(* IEC 61131-3 sources: TetherPLC/compat/tc2 (part 5) *)

(* ---- tc2_nci.st ---- *)
// Tc2_NCI — TwinCAT NC-I (TF5100) channel-interpolation surface over
// the builtin FB_MotionAxis (tplc-motion service). This file
// implements the interpolation core: coordinated multi-axis
// setpoint streaming in CyclicSyncPosition (CSP, mode 8).
//
// Model: TwinCAT's NC-I runs a G-code / FIFO interpreter in the NC
// kernel that emits per-axis position setpoints every NC cycle to
// axes in CSP mode. The compat model collapses one in-flight
// geometric block into each FB: FB_NciLine parameterizes a straight
// line across a 3-axis group, advances the path parameter s by
// Velocity*CycleUs each scan, and streams per-axis targets
// (0x607A) with the axes in CSP mode — which is exactly how the NC
// kernel drives CSP axes. There is no backend group registry, so a
// "3D group" is just the X/Y/Z axis handles passed to the block
// (TwinCAT's CfgBuild3DGroup maps to passing those handles).
//
// Time base: the FB has no access to the host clock, so the caller
// supplies the scan period via CycleUs (microseconds); path
// Velocity is then in user-units/second and s += Velocity*CycleUs/1e6
// per scan. Positions/velocities are the backend's int32 user
// units (TwinCAT LREAL — documented gap). Determinism: under --sim,
// CycleUs = step_us makes the path advance a fixed amount per step,
// and CSP snaps each axis to the streamed target so commanded and
// actual positions match.
//
// G-code interpretation lives in Tether: tether_io_motion_server
// exposes an nc.* channel that compiles program text with its G-code
// interpreter, time-parameterizes it with the motion planner (corner
// blending, jerk-limited profiles), and streams CSP setpoints to the
// drives on the mc.time clock. The FB_NciChan blocks below are the
// PLC-side control surface for that channel (TwinCAT Itp* shape);
// there is no in-process interpreter — with no TPLC_MOTION_IO
// endpoint the blocks report the service as unavailable.
//
// Honest gaps: FB_NciLine is the foundational interpreter-free path
// (single block, no queue); the nc.* channel has no PLC-visible
// M-function handshake, R-parameters, zero-shift, or cyclic-channel
// offset tables yet. See DECISIONS D-IMPL-56.
// SPDX-License-Identifier: Apache-2.0 OR MPL-2.0

// ---- F_NciSqrt: Newton (Babylonian) square root for LREAL ----
// The ST layer has no SQRT builtin, so the path length is computed
// with a fixed-iteration Newton iteration. r0 = x/2 + 1 converges
// monotonically for x >= 0; 48 iterations is enough for the full
// int32 path range and keeps the result deterministic.
FUNCTION F_NciSqrt : LREAL
VAR_INPUT
    x : LREAL;
END_VAR
VAR
    r : LREAL;
    k : INT;
END_VAR
    IF x <= 0.0 THEN
        F_NciSqrt := 0.0;
    ELSE
        r := x * 0.5 + 1.0;
        k := 0;
        REPEAT
            r := 0.5 * (r + x / r);
            k := k + 1;
        UNTIL k >= 48
        END_REPEAT;
        F_NciSqrt := r;
    END_IF;
END_FUNCTION

// ---- FB_NciLine: coordinated 3-axis linear move (CSP stream) ----
// On Execute, latches each axis's actual position as the segment
// start, computes deltas and the Euclidean path length, switches
// all three axes to CSP mode, then each scan advances s toward len
// and writes each axis's interpolated TargetPosition. Done when
// s reaches len (all axes arrive simultaneously — a straight line).
// Releasing Execute mid-move aborts: streaming stops, so each axis
// holds its last streamed target (CommandAborted pulses).
FUNCTION_BLOCK FB_NciLine
VAR_INPUT
    Execute : BOOL;
    PosX : DINT;
    PosY : DINT;
    PosZ : DINT;
    Velocity : DINT;    // resultant path velocity, user-units/sec
    CycleUs : DINT;     // scan period, microseconds
    AxisX : UDINT;
    AxisY : UDINT;
    AxisZ : UDINT;
END_VAR
VAR_OUTPUT
    Done : BOOL;
    Busy : BOOL;
    CommandAborted : BOOL;
    Error : BOOL;
    ErrorID : UDINT;
    ActPosX : DINT;     // interpolated commanded positions
    ActPosY : DINT;
    ActPosZ : DINT;
    PathLen : DINT;     // Euclidean path length (user units)
    PathS : DINT;       // current path parameter along the line
END_VAR
VAR
    axX : FB_MotionAxis;
    axY : FB_MotionAxis;
    axZ : FB_MotionAxis;
    exPrev : BOOL;
    exEdge : BOOL;
    active : BOOL;
    sxr : LREAL;
    syr : LREAL;
    szr : LREAL;
    dxr : LREAL;
    dyr : LREAL;
    dzr : LREAL;
    len : LREAL;
    s : LREAL;
    dt : LREAL;
    vel : LREAL;
END_VAR
    // advance every axis's dynamics once per scan (one poll advances
    // the whole pool); bind each instance to its group axis
    axX.OP := 3; axX();
    axX.AXIS := AxisX; axY.AXIS := AxisY; axZ.AXIS := AxisZ;
    exEdge := Execute AND NOT exPrev;
    exPrev := Execute;
    Done := FALSE;
    CommandAborted := FALSE;
    Error := FALSE;
    ErrorID := 0;

    IF exEdge THEN
        // latch the segment start = current actual positions
        axX.OP := 4; axX.INDEX := 16#6064; axX();
        sxr := DINT_TO_LREAL(axX.VALUE);
        axY.OP := 4; axY.INDEX := 16#6064; axY();
        syr := DINT_TO_LREAL(axY.VALUE);
        axZ.OP := 4; axZ.INDEX := 16#6064; axZ();
        szr := DINT_TO_LREAL(axZ.VALUE);
        dxr := DINT_TO_LREAL(PosX) - sxr;
        dyr := DINT_TO_LREAL(PosY) - syr;
        dzr := DINT_TO_LREAL(PosZ) - szr;
        len := F_NciSqrt(dxr * dxr + dyr * dyr + dzr * dzr);
        PathLen := TRUNC(len);
        dt := DINT_TO_LREAL(CycleUs) / 1000000.0;
        vel := DINT_TO_LREAL(Velocity);
        s := 0.0;
        IF len < 0.5 THEN
            // already at the target — nothing to stream
            active := FALSE;
            Done := TRUE;
        ELSE
            // put the group into CyclicSyncPosition (mode 8)
            axX.OP := 5; axX.INDEX := 16#6060; axX.VALUE := 8; axX();
            axY.OP := 5; axY.INDEX := 16#6060; axY.VALUE := 8; axY();
            axZ.OP := 5; axZ.INDEX := 16#6060; axZ.VALUE := 8; axZ();
            active := TRUE;
        END_IF;
    END_IF;

    IF active THEN
        IF Execute THEN
            // advance the path parameter and clamp at the end
            s := s + vel * dt;
            IF s >= len THEN
                s := len;
                active := FALSE;
                Done := TRUE;
            END_IF;
            PathS := TRUNC(s);
            // stream the interpolated setpoints to each CSP axis
            ActPosX := TRUNC(sxr + dxr * s / len);
            ActPosY := TRUNC(syr + dyr * s / len);
            ActPosZ := TRUNC(szr + dzr * s / len);
            axX.OP := 5; axX.INDEX := 16#607A; axX.VALUE := ActPosX; axX();
            axY.OP := 5; axY.INDEX := 16#607A; axY.VALUE := ActPosY; axY();
            axZ.OP := 5; axZ.INDEX := 16#607A; axZ.VALUE := ActPosZ; axZ();
        ELSE
            // aborted: stop streaming so each axis holds its last
            // CSP setpoint (position freezes in place)
            active := FALSE;
            CommandAborted := TRUE;
        END_IF;
    END_IF;
    Busy := active;
END_FUNCTION_BLOCK

// ---- FB_NciEStop: cut power to a 3-axis group ----
// On Execute it writes DisableVoltage (controlword 0x0000) to each
// axis so the group coasts to a stop; Status reports all three
// axes left OperationEnabled. Honest E-stop: a real NC fault also
// freezes the interpolator, which the caller models by releasing
// FB_NciLine's Execute.
FUNCTION_BLOCK FB_NciEStop
VAR_INPUT
    Execute : BOOL;
    AxisX : UDINT;
    AxisY : UDINT;
    AxisZ : UDINT;
END_VAR
VAR_OUTPUT
    Status : BOOL;
    Busy : BOOL;
    Error : BOOL;
    ErrorID : UDINT;
END_VAR
VAR
    ax : FB_MotionAxis;
    exPrev : BOOL;
    exEdge : BOOL;
END_VAR
    ax.OP := 3; ax();
    exEdge := Execute AND NOT exPrev;
    exPrev := Execute;
    Error := FALSE;
    ErrorID := 0;
    IF exEdge THEN
        ax.AXIS := AxisX; ax.OP := 5; ax.INDEX := 16#6040; ax.VALUE := 0; ax();
        ax.AXIS := AxisY; ax.OP := 5; ax.INDEX := 16#6040; ax.VALUE := 0; ax();
        ax.AXIS := AxisZ; ax.OP := 5; ax.INDEX := 16#6040; ax.VALUE := 0; ax();
    END_IF;
    // Status = all three axes out of OperationEnabled (state <> 39)
    ax.AXIS := AxisX; ax.OP := 6; ax();
    Status := (ax.STATUS <> 39);
    ax.AXIS := AxisY; ax.OP := 6; ax();
    Status := Status AND (ax.STATUS <> 39);
    ax.AXIS := AxisZ; ax.OP := 6; ax();
    Status := Status AND (ax.STATUS <> 39);
    Busy := Execute AND NOT Status;
END_FUNCTION_BLOCK

// ---- NC interpreter channel (Tether-owned G-code) ----
// Command codes written to FB_NciChan.CMD (nc.cmd on the wire):
//   1=run 2=step 3=pause 4=resume 5=stop 6=reset 7=verify
// Channel states reported by FB_NciChan.STATE (nc.state):
//   0=idle 1=ready 2=running 3=paused 4=finished 5=error 6=stopped

// ---- FB_ItpLoadText: upload inline program text to the channel ----
// Rising edge on Execute writes PROG to nc.prog; the server compiles
// it immediately. Done means the text was accepted (compile status is
// visible via FB_ItpStatus/nc.state afterwards). TwinCAT loads files
// through ItpLoadProg; inline text is the Tether-native path.
FUNCTION_BLOCK FB_ItpLoadText
VAR_INPUT
    Execute : BOOL;
    ChanId : UDINT;
    ProgText : STRING[4095];
END_VAR
VAR_OUTPUT
    Done : BOOL;
    Busy : BOOL;
    Error : BOOL;
    ErrorID : UDINT;
END_VAR
VAR
    ch : FB_NciChan;
    exPrev : BOOL;
END_VAR
    Done := FALSE;
    Error := FALSE;
    ErrorID := 0;
    IF Execute AND NOT exPrev THEN
        ch.OP := 1;
        ch.CHAN := ChanId;
        ch.PROG := ProgText;
        ch();
        IF ch.STATUS = 0 THEN
            Done := TRUE;
        ELSE
            Error := TRUE;
            ErrorID := ch.ERRID;
        END_IF;
    END_IF;
    exPrev := Execute;
    Busy := FALSE;
END_FUNCTION_BLOCK

// ---- FB_ItpLoadProg: load a program file on the server host ----
// Rising edge on Execute writes PathName to nc.prog_path; the server
// opens and compiles the file. Mirrors TwinCAT ItpLoadProg(Ex).
FUNCTION_BLOCK FB_ItpLoadProg
VAR_INPUT
    Execute : BOOL;
    ChanId : UDINT;
    PathName : STRING[127];
END_VAR
VAR_OUTPUT
    Done : BOOL;
    Busy : BOOL;
    Error : BOOL;
    ErrorID : UDINT;
END_VAR
VAR
    ch : FB_NciChan;
    exPrev : BOOL;
END_VAR
    Done := FALSE;
    Error := FALSE;
    ErrorID := 0;
    IF Execute AND NOT exPrev THEN
        ch.OP := 2;
        ch.CHAN := ChanId;
        ch.PATH := PathName;
        ch();
        IF ch.STATUS = 0 THEN
            Done := TRUE;
        ELSE
            Error := TRUE;
            ErrorID := ch.ERRID;
        END_IF;
    END_IF;
    exPrev := Execute;
    Busy := FALSE;
END_FUNCTION_BLOCK

// ---- FB_ItpStartStop: start/stop the NC channel ----
// Rising edge on Start issues cmd RUN, on Stop issues cmd STOP.
// Mirrors TwinCAT ItpStartStopEx (bStart/bStop).
FUNCTION_BLOCK FB_ItpStartStop
VAR_INPUT
    Start : BOOL;
    Stop : BOOL;
    ChanId : UDINT;
END_VAR
VAR_OUTPUT
    Done : BOOL;
    Busy : BOOL;
    Error : BOOL;
    ErrorID : UDINT;
END_VAR
VAR
    ch : FB_NciChan;
    stPrev : BOOL;
    spPrev : BOOL;
END_VAR
    Done := FALSE;
    Error := FALSE;
    ErrorID := 0;
    IF Start AND NOT stPrev THEN
        ch.OP := 3;
        ch.CHAN := ChanId;
        ch.CMD := 1;
        ch();
        IF ch.STATUS = 0 THEN
            Done := TRUE;
        ELSE
            Error := TRUE;
            ErrorID := ch.ERRID;
        END_IF;
    END_IF;
    IF Stop AND NOT spPrev THEN
        ch.OP := 3;
        ch.CHAN := ChanId;
        ch.CMD := 5;
        ch();
        IF ch.STATUS = 0 THEN
            Done := TRUE;
        ELSE
            Error := TRUE;
            ErrorID := ch.ERRID;
        END_IF;
    END_IF;
    stPrev := Start;
    spPrev := Stop;
    Busy := FALSE;
END_FUNCTION_BLOCK

// ---- FB_ItpReset: reset the NC channel ----
// Rising edge issues cmd RESET: clears program, state and errors.
// Mirrors TwinCAT ItpResetEx.
FUNCTION_BLOCK FB_ItpReset
VAR_INPUT
    Execute : BOOL;
    ChanId : UDINT;
END_VAR
VAR_OUTPUT
    Done : BOOL;
    Busy : BOOL;
    Error : BOOL;
    ErrorID : UDINT;
END_VAR
VAR
    ch : FB_NciChan;
    exPrev : BOOL;
END_VAR
    Done := FALSE;
    Error := FALSE;
    ErrorID := 0;
    IF Execute AND NOT exPrev THEN
        ch.OP := 3;
        ch.CHAN := ChanId;
        ch.CMD := 6;
        ch();
        IF ch.STATUS = 0 THEN
            Done := TRUE;
        ELSE
            Error := TRUE;
            ErrorID := ch.ERRID;
        END_IF;
    END_IF;
    exPrev := Execute;
    Busy := FALSE;
END_FUNCTION_BLOCK

// ---- FB_ItpEStop: emergency stop on the channel ----
// Rising edge issues cmd STOP: the channel drops out of RUNNING and
// the planner holds the last setpoints (the sim axes freeze). A
// machine E-stop also cuts axis power — compose with FB_NciEStop
// for that. Mirrors TwinCAT ItpEStopEx.
FUNCTION_BLOCK FB_ItpEStop
VAR_INPUT
    Execute : BOOL;
    ChanId : UDINT;
END_VAR
VAR_OUTPUT
    Done : BOOL;
    Busy : BOOL;
    Error : BOOL;
    ErrorID : UDINT;
END_VAR
VAR
    ch : FB_NciChan;
    exPrev : BOOL;
END_VAR
    Done := FALSE;
    Error := FALSE;
    ErrorID := 0;
    IF Execute AND NOT exPrev THEN
        ch.OP := 3;
        ch.CHAN := ChanId;
        ch.CMD := 5;
        ch();
        IF ch.STATUS = 0 THEN
            Done := TRUE;
        ELSE
            Error := TRUE;
            ErrorID := ch.ERRID;
        END_IF;
    END_IF;
    exPrev := Execute;
    Busy := FALSE;
END_FUNCTION_BLOCK

// ---- FB_ItpStatus: cyclic channel status ----
// Polls nc.state/line/total/errcode/progress/duration every scan and
// mirrors them to the outputs (call unconditionally each cycle).
// Finished is TRUE in FINISHED/ERROR/STOPPED; IsEStop is TRUE when
// the channel is in STOPPED, matching TwinCAT ItpIsEStop semantics.
FUNCTION_BLOCK FB_ItpStatus
VAR_INPUT
    ChanId : UDINT;
END_VAR
VAR_OUTPUT
    Valid : BOOL;
    State : DINT;
    Line : UDINT;
    Total : UDINT;
    ErrCode : DINT;
    Finished : BOOL;
    IsEStop : BOOL;
    ProgressMs : DINT;
    DurationMs : DINT;
    MFunc : UDINT;
    FifoLen : UDINT;
    FifoSeq : UDINT;
    Error : BOOL;
    ErrorID : UDINT;
END_VAR
VAR
    ch : FB_NciChan;
END_VAR
    ch.OP := 4;
    ch.CHAN := ChanId;
    ch();
    Valid := (ch.STATUS = 0);
    Error := NOT Valid;
    ErrorID := ch.ERRID;
    State := 0;
    Line := 0;
    Total := 0;
    ErrCode := 0;
    Finished := FALSE;
    IsEStop := FALSE;
    ProgressMs := 0;
    DurationMs := 0;
    IF Valid THEN
        State := ch.STATE;
        Line := ch.LINE;
        Total := ch.TOTAL;
        ErrCode := ch.NERR;
        Finished := (State = 4) OR (State = 5) OR (State = 6);
        IsEStop := (State = 6);
        ProgressMs := ch.PROGRESS;
        DurationMs := ch.DURATION;
        MFunc := ch.MFUNC;
        FifoLen := ch.FIFOLEN;
        FifoSeq := ch.FIFOSEQ;
    END_IF;
END_FUNCTION_BLOCK

// ---- FB_ItpFiFoWrite: append a block to the channel FIFO queue ----
// Rising edge on Execute writes Block (one G-code block) to nc.fifo;
// queued entries execute in order after the active plan, anchored at
// the last commanded position. Mirrors TwinCAT FiFoWrite semantics.
FUNCTION_BLOCK FB_ItpFiFoWrite
VAR_INPUT
    Execute : BOOL;
    ChanId : UDINT;
    Block : STRING[127];
END_VAR
VAR_OUTPUT
    Done : BOOL;
    Busy : BOOL;
    Error : BOOL;
    ErrorID : UDINT;
END_VAR
VAR
    ch : FB_NciChan;
    exPrev : BOOL;
END_VAR
    Done := FALSE;
    Error := FALSE;
    ErrorID := 0;
    IF Execute AND NOT exPrev THEN
        ch.OP := 5;
        ch.CHAN := ChanId;
        ch.PROG := Block;
        ch();
        IF ch.STATUS = 0 THEN
            Done := TRUE;
        ELSE
            Error := TRUE;
            ErrorID := ch.ERRID;
        END_IF;
    END_IF;
    exPrev := Execute;
    Busy := FALSE;
END_FUNCTION_BLOCK

// ---- FB_ItpConfirmHsk: confirm a pending M-function ----
// Rising edge confirms the M-code reported in sts.MFunc; the held
// channel resumes. Mirrors TwinCAT ItpConfirmHsk.
FUNCTION_BLOCK FB_ItpConfirmHsk
VAR_INPUT
    Execute : BOOL;
    ChanId : UDINT;
END_VAR
VAR_OUTPUT
    Done : BOOL;
    Busy : BOOL;
    Error : BOOL;
    ErrorID : UDINT;
END_VAR
VAR
    ch : FB_NciChan;
    exPrev : BOOL;
END_VAR
    Done := FALSE;
    Error := FALSE;
    ErrorID := 0;
    IF Execute AND NOT exPrev THEN
        ch.OP := 6;
        ch.CHAN := ChanId;
        ch();
        IF ch.STATUS = 0 THEN
            Done := TRUE;
        ELSE
            Error := TRUE;
            ErrorID := ch.ERRID;
        END_IF;
    END_IF;
    exPrev := Execute;
    Busy := FALSE;
END_FUNCTION_BLOCK

// ---- FB_ItpWriteRParam: write one R-parameter register ----
// Rising edge stores Value into R-parameter Index on the channel;
// applied on the next program compile. Mirrors ItpWriteRParams.
FUNCTION_BLOCK FB_ItpWriteRParam
VAR_INPUT
    Execute : BOOL;
    ChanId : UDINT;
    Index : UDINT;
    Value : LREAL;
END_VAR
VAR_OUTPUT
    Done : BOOL;
    Busy : BOOL;
    Error : BOOL;
    ErrorID : UDINT;
END_VAR
VAR
    ch : FB_NciChan;
    exPrev : BOOL;
END_VAR
    Done := FALSE;
    Error := FALSE;
    ErrorID := 0;
    IF Execute AND NOT exPrev THEN
        ch.OP := 7;
        ch.CHAN := ChanId;
        ch.AUX := Index;
        ch.RVAL := Value;
        ch();
        IF ch.STATUS = 0 THEN
            Done := TRUE;
        ELSE
            Error := TRUE;
            ErrorID := ch.ERRID;
        END_IF;
    END_IF;
    exPrev := Execute;
    Busy := FALSE;
END_FUNCTION_BLOCK

// ---- FB_ItpReadRParam: read one R-parameter register ----
// Rising edge reads R-parameter Index into Value. Mirrors
// ItpReadRParams.
FUNCTION_BLOCK FB_ItpReadRParam
VAR_INPUT
    Execute : BOOL;
    ChanId : UDINT;
    Index : UDINT;
END_VAR
VAR_OUTPUT
    Done : BOOL;
    Busy : BOOL;
    Error : BOOL;
    ErrorID : UDINT;
    Value : LREAL;
END_VAR
VAR
    ch : FB_NciChan;
    exPrev : BOOL;
END_VAR
    Done := FALSE;
    Error := FALSE;
    ErrorID := 0;
    IF Execute AND NOT exPrev THEN
        ch.OP := 8;
        ch.CHAN := ChanId;
        ch.AUX := Index;
        ch();
        IF ch.STATUS = 0 THEN
            Done := TRUE;
            Value := ch.RVAL;
        ELSE
            Error := TRUE;
            ErrorID := ch.ERRID;
        END_IF;
    END_IF;
    exPrev := Execute;
    Busy := FALSE;
END_FUNCTION_BLOCK

// ---- FB_ItpZeroShift: write the channel zero-shift offsets ----
// Rising edge stores the XYZ offsets; applied as a G92 prefix on the
// next program compile.
FUNCTION_BLOCK FB_ItpZeroShift
VAR_INPUT
    Execute : BOOL;
    ChanId : UDINT;
    OffX : LREAL;
    OffY : LREAL;
    OffZ : LREAL;
END_VAR
VAR_OUTPUT
    Done : BOOL;
    Busy : BOOL;
    Error : BOOL;
    ErrorID : UDINT;
END_VAR
VAR
    ch : FB_NciChan;
    exPrev : BOOL;
END_VAR
    Done := FALSE;
    Error := FALSE;
    ErrorID := 0;
    IF Execute AND NOT exPrev THEN
        ch.OP := 9;
        ch.CHAN := ChanId;
        ch.ZSX := OffX;
        ch.ZSY := OffY;
        ch.ZSZ := OffZ;
        ch();
        IF ch.STATUS = 0 THEN
            Done := TRUE;
        ELSE
            Error := TRUE;
            ErrorID := ch.ERRID;
        END_IF;
    END_IF;
    exPrev := Execute;
    Busy := FALSE;
END_FUNCTION_BLOCK

(* ---- tc2_nckin.st ---- *)
// tc2_nckin.st — Tc2_NcKinematicTransformation: kinematic
// transformation objects (12 APIs) over the tplc-kin service /
// FB_Kin builtin. The transform engine is the Tether kinematics
// library (ForwardKinematics.hpp): forward maps joint values to a
// Pose6D, backward runs deterministic damped least-squares position
// IK (orientation unconstrained, max 8 DOF).
//
// Object model: up to 8 transformation objects (oidTrafo 0..7),
// each with a configured chain type (cartesian, planar2d,
// articulated3, scara, serial6, serial7, gantry5, delta, stewart),
// optional ACS (joint) and MCS (Cartesian) axis lists, a parameter
// lock, a rotation preset, and an NC channel id. Chain geometry is
// configured through FB_Kin directly (OP1) or the compat case; the
// TwinCAT project-side configuration surface is flattened into the
// oidTrafo object index.
//
// Flattening vs the TwinCAT signatures:
//   ST_KinAxes          -> AcsAxis/McsAxis : ARRAY[0..7] OF UDINT
//                          (axis handles, 0 = empty slot; the
//                          configured count is the leading run of
//                          non-zero entries)
//   NCTOPLC_NCICHANNEL_REF -> nItpChannelId : UDINT
//   U_KinMetaInfo       -> oidTrafo input (object id) + MetaState /
//                          MetaError outputs
//   oidTrafo on blocks  -> kinematic object index 0..7 (TwinCAT
//                          binds the object via the project)
//   pDataIn/pDataOut    -> InData/OutData : ARRAY[0..7] OF LREAL +
//                          nSizeIn/nSizeOut element counts (the
//                          byte-pointer contract is flattened)
//   stAxesPosIn/Out     -> VAR_IN_OUT ARRAY[0..7] OF LREAL
//   stRotation          -> Rotation : ARRAY[0..2] OF LREAL
//   E_KINSTATUS         -> UDINT (0 idle 1 ready 2 error 3 homing)
//   FUNCTIONs with output params -> FUNCTION_BLOCKs (dialect rule)
//
// FB_Kin OP map: 1 configure, 2 set axes, 3 command, 4 calc input,
// 5 result, 6 set locked, 7 rotation, 8 status, 9 set channel,
// 10 get axes.

// Shared pump: run one FB_Kin op sequence on the rising edge.
FUNCTION_BLOCK KinPump
VAR_INPUT
    OP      : UDINT;
    OBJ     : UDINT;
    TYPE_   : DINT;
    PRESET  : UDINT;
    NCFG    : UDINT;
    NIN     : UDINT;
    NACS    : UDINT;
    NMCS    : UDINT;
    CMD     : UDINT;
    ROP     : UDINT;
    CHN     : UDINT;
    LOCKED  : UDINT;
    bExecute : BOOL;
END_VAR
VAR_OUTPUT
    bBusy   : BOOL;
    bError  : BOOL;
    nErrorId : UDINT;
END_VAR
VAR
    kin : FB_Kin;
    exPrev : BOOL;
    i : UDINT;
END_VAR
    bBusy := FALSE;
    bError := FALSE;
    nErrorId := 0;
    IF bExecute AND NOT exPrev THEN
        bBusy := TRUE;
        kin.OBJ := OBJ;
        kin.OP := OP;
        kin.TYPEIN := TYPE_;
        kin.PRESET := PRESET;
        kin.NCFG := NCFG;
        kin.NIN := NIN;
        kin.NACS := NACS;
        kin.NMCS := NMCS;
        kin.CMD := CMD;
        kin.ROP := ROP;
        kin.CHN := CHN;
        kin.LOCKED := LOCKED;
        FOR i := 0 TO 31 DO
            kin.CFG[i] := 0.0;
        END_FOR;
        kin();
        IF kin.STATUS <> 0 THEN
            bError := TRUE;
            nErrorId := kin.ERRID;
        END_IF;
    END_IF;
    exPrev := bExecute;
END_FUNCTION_BLOCK

// ---- FB_KinConfigGroup: bind ACS/MCS axes + channel to object ----
FUNCTION_BLOCK FB_KinConfigGroup
VAR_INPUT
    bExecute : BOOL;
    bCartesianMode : BOOL;
    oidTrafo : UDINT;
    nItpChannelId : UDINT;
    AcsAxis : ARRAY[0..7] OF UDINT;
    McsAxis : ARRAY[0..7] OF UDINT;
END_VAR
VAR_OUTPUT
    bBusy : BOOL;
    bError : BOOL;
    nErrorId : UDINT;
END_VAR
VAR
    kin : FB_Kin;
    exPrev : BOOL;
    i : UDINT;
    nAcs : UDINT;
    nMcs : UDINT;
END_VAR
    bBusy := FALSE;
    bError := FALSE;
    nErrorId := 0;
    IF bExecute AND NOT exPrev THEN
        bBusy := TRUE;
        /* count the leading run of non-zero (1-based) handles */
        nAcs := 0;
        FOR i := 0 TO 7 DO
            IF AcsAxis[i] <> 0 AND i = nAcs THEN
                nAcs := nAcs + 1;
            END_IF;
        END_FOR;
        nMcs := 0;
        FOR i := 0 TO 7 DO
            IF McsAxis[i] <> 0 AND i = nMcs THEN
                nMcs := nMcs + 1;
            END_IF;
        END_FOR;
        kin.OBJ := oidTrafo;
        kin.OP := 2;
        kin.NACS := nAcs;
        kin.NMCS := nMcs;
        FOR i := 0 TO 7 DO
            kin.ACS[i] := 0;
            kin.MCS[i] := 0;
        END_FOR;
        IF nAcs > 0 THEN
            FOR i := 0 TO nAcs - 1 DO
                kin.ACS[i] := AcsAxis[i];
            END_FOR;
        END_IF;
        IF nMcs > 0 THEN
            FOR i := 0 TO nMcs - 1 DO
                kin.MCS[i] := McsAxis[i];
            END_FOR;
        END_IF;
        kin();
        IF kin.STATUS <> 0 THEN
            bError := TRUE;
            nErrorId := kin.ERRID;
        ELSE
            kin.OP := 9;
            kin.CHN := nItpChannelId;
            kin();
            IF kin.STATUS <> 0 THEN
                bError := TRUE;
                nErrorId := kin.ERRID;
            END_IF;
        END_IF;
    END_IF;
    exPrev := bExecute;
END_FUNCTION_BLOCK

// ---- FB_KinResetGroup: reset the kinematic group ----
FUNCTION_BLOCK FB_KinResetGroup
VAR_INPUT
    bExecute : BOOL;
    oidTrafo : UDINT;
    nItpChannelId : UDINT;
END_VAR
VAR_OUTPUT
    bBusy : BOOL;
    bError : BOOL;
    nErrorId : UDINT;
END_VAR
VAR
    kin : FB_Kin;
    exPrev : BOOL;
END_VAR
    bBusy := FALSE;
    bError := FALSE;
    nErrorId := 0;
    IF bExecute AND NOT exPrev THEN
        bBusy := TRUE;
        kin.OBJ := oidTrafo;
        kin.OP := 3;
        kin.CMD := 3;   /* TPLC_KIN_CMD_RESET */
        kin();
        IF kin.STATUS <> 0 THEN
            bError := TRUE;
            nErrorId := kin.ERRID;
        END_IF;
        /* re-associate the channel when one is given */
        IF nItpChannelId <> 0 AND NOT bError THEN
            kin.OP := 9;
            kin.CHN := nItpChannelId;
            kin();
            IF kin.STATUS <> 0 THEN
                bError := TRUE;
                nErrorId := kin.ERRID;
            END_IF;
        END_IF;
    END_IF;
    exPrev := bExecute;
END_FUNCTION_BLOCK

// ---- FB_KinCalcTrafo: forward / backward transform ----
FUNCTION_BLOCK FB_KinCalcTrafo
VAR_INPUT
    bExecute : BOOL;
    bForward : BOOL;
    oidTrafo : UDINT;
END_VAR
VAR_IN_OUT
    AxesPosIn : ARRAY[0..7] OF LREAL;
    AxesPosOut : ARRAY[0..7] OF LREAL;
    MetaState : UDINT;
    MetaError : UDINT;
END_VAR
VAR_OUTPUT
    bBusy : BOOL;
    bError : BOOL;
    nErrorId : UDINT;
END_VAR
VAR
    kin : FB_Kin;
    exPrev : BOOL;
    i : UDINT;
    cmd : UDINT;
END_VAR
    bBusy := FALSE;
    bError := FALSE;
    nErrorId := 0;
    MetaState := 0;
    MetaError := 0;
    IF bExecute AND NOT exPrev THEN
        bBusy := TRUE;
        kin.OBJ := oidTrafo;
        /* input: forward = joints, backward = target xyz + seed */
        kin.OP := 4;
        kin.NIN := 8;
        FOR i := 0 TO 7 DO
            kin.IN[i] := AxesPosIn[i];
        END_FOR;
        kin();
        IF kin.STATUS <> 0 THEN
            bError := TRUE;
            nErrorId := kin.ERRID;
        ELSE
            cmd := 2;   /* backward (IK) */
            IF bForward THEN cmd := 1; END_IF;
            kin.OP := 3;
            kin.CMD := cmd;
            kin();
            IF kin.STATUS <> 0 THEN
                bError := TRUE;
                nErrorId := kin.ERRID;
            ELSE
                kin.OP := 5;
                kin();
                IF kin.STATUS <> 0 THEN
                    bError := TRUE;
                    nErrorId := kin.ERRID;
                ELSE
                    /* ERR/STATE only refresh on OP8; poll once so
                       MetaError carries the object's error code
                       (e.g. 1 = no model, 3 = IK no convergence). */
                    kin.OP := 8;
                    kin();
                    MetaState := kin.STATE;
                    MetaError := kin.ERR;
                    IF bForward THEN
                        /* pose x,y,z,roll,pitch,yaw -> out[0..5] */
                        FOR i := 0 TO 5 DO
                            AxesPosOut[i] := kin.OUT[i];
                        END_FOR;
                    ELSE
                        /* IK joint solution q -> out[0..7] */
                        FOR i := 0 TO 7 DO
                            AxesPosOut[i] := kin.Q[i];
                        END_FOR;
                    END_IF;
                END_IF;
            END_IF;
        END_IF;
    END_IF;
    exPrev := bExecute;
END_FUNCTION_BLOCK

// ---- FB_KinCalcMultiTrafo: flattened single-object transform ----
// TwinCAT packs a caller buffer of transform requests; the flattened
// form carries one object's input vector and returns the result
// vector (pose for forward, joints for backward).
FUNCTION_BLOCK FB_KinCalcMultiTrafo
VAR_INPUT
    bExecute : BOOL;
    bForward : BOOL;
    oidTrafo : UDINT;
    nSizeIn : UDINT;
    nSizeOut : UDINT;
END_VAR
VAR_IN_OUT
    InData : ARRAY[0..7] OF LREAL;
    OutData : ARRAY[0..15] OF LREAL;
END_VAR
VAR_OUTPUT
    bBusy : BOOL;
    bError : BOOL;
    nErrorId : UDINT;
    nOutLen : UDINT;
END_VAR
VAR
    kin : FB_Kin;
    exPrev : BOOL;
    i : UDINT;
    n : UDINT;
    cmd : UDINT;
END_VAR
    bBusy := FALSE;
    bError := FALSE;
    nErrorId := 0;
    nOutLen := 0;
    IF bExecute AND NOT exPrev THEN
        bBusy := TRUE;
        kin.OBJ := oidTrafo;
        n := nSizeIn;
        IF n > 8 THEN n := 8; END_IF;
        kin.OP := 4;
        kin.NIN := n;
        FOR i := 0 TO 7 DO
            kin.IN[i] := 0.0;
        END_FOR;
        IF n > 0 THEN
            FOR i := 0 TO n - 1 DO
                kin.IN[i] := InData[i];
            END_FOR;
        END_IF;
        kin();
        IF kin.STATUS <> 0 THEN
            bError := TRUE;
            nErrorId := kin.ERRID;
        ELSE
            cmd := 2;
            IF bForward THEN cmd := 1; END_IF;
            kin.OP := 3;
            kin.CMD := cmd;
            kin();
            IF kin.STATUS <> 0 THEN
                bError := TRUE;
                nErrorId := kin.ERRID;
            ELSE
                kin.OP := 5;
                kin();
                IF kin.STATUS <> 0 THEN
                    bError := TRUE;
                    nErrorId := kin.ERRID;
                ELSE
                    IF bForward THEN
                        FOR i := 0 TO 7 DO
                            OutData[i] := kin.OUT[i];
                        END_FOR;
                    ELSE
                        FOR i := 0 TO 7 DO
                            OutData[i] := kin.Q[i];
                        END_FOR;
                    END_IF;
                    nOutLen := 8;
                END_IF;
            END_IF;
        END_IF;
    END_IF;
    exPrev := bExecute;
END_FUNCTION_BLOCK

// ---- FB_KinUnlockTrafoParam / FB_KinLockTrafoParam ----
FUNCTION_BLOCK FB_KinUnlockTrafoParam
VAR_INPUT
    bExecute : BOOL;
    oidTrafo : UDINT;
END_VAR
VAR_OUTPUT
    bBusy : BOOL;
    bError : BOOL;
    nErrorId : UDINT;
END_VAR
VAR
    p : KinPump;
END_VAR
    p.OP := 6; p.OBJ := oidTrafo; p.LOCKED := 0;
    p.bExecute := bExecute;
    p();
    bBusy := p.bBusy; bError := p.bError; nErrorId := p.nErrorId;
END_FUNCTION_BLOCK

FUNCTION_BLOCK FB_KinLockTrafoParam
VAR_INPUT
    bExecute : BOOL;
    oidTrafo : UDINT;
END_VAR
VAR_OUTPUT
    bBusy : BOOL;
    bError : BOOL;
    nErrorId : UDINT;
END_VAR
VAR
    p : KinPump;
END_VAR
    p.OP := 6; p.OBJ := oidTrafo; p.LOCKED := 1;
    p.bExecute := bExecute;
    p();
    bBusy := p.bBusy; bError := p.bError; nErrorId := p.nErrorId;
END_FUNCTION_BLOCK

// ---- FB_KinExtendedRotationRange: save on execute edge, restore
// on release (extends the achievable rotation range temporarily).
FUNCTION_BLOCK FB_KinExtendedRotationRange
VAR_INPUT
    bExecute : BOOL;
    oidTrafo : UDINT;
END_VAR
VAR_OUTPUT
    bBusy : BOOL;
    bError : BOOL;
    nErrorId : UDINT;
END_VAR
VAR
    kin : FB_Kin;
    exPrev : BOOL;
    rop : UDINT;
END_VAR
    bBusy := FALSE;
    bError := FALSE;
    nErrorId := 0;
    rop := 0;
    IF bExecute AND NOT exPrev THEN
        rop := 2;   /* TPLC_KIN_ROT_SAVE */
        bBusy := TRUE;
    ELSIF NOT bExecute AND exPrev THEN
        rop := 3;   /* TPLC_KIN_ROT_RESTORE */
        bBusy := TRUE;
    END_IF;
    IF rop <> 0 THEN
        kin.OBJ := oidTrafo;
        kin.OP := 7;
        kin.ROP := rop;
        kin();
        IF kin.STATUS <> 0 THEN
            bError := TRUE;
            nErrorId := kin.ERRID;
        END_IF;
    END_IF;
    exPrev := bExecute;
END_FUNCTION_BLOCK

// ---- FB_KinPresetRotation: set the rotational state ----
FUNCTION_BLOCK FB_KinPresetRotation
VAR_INPUT
    bExecute : BOOL;
    oidTrafo : UDINT;
END_VAR
VAR_IN_OUT
    Rotation : ARRAY[0..2] OF LREAL;
END_VAR
VAR_OUTPUT
    bBusy : BOOL;
    bError : BOOL;
    nErrorId : UDINT;
END_VAR
VAR
    kin : FB_Kin;
    exPrev : BOOL;
    i : UDINT;
END_VAR
    bBusy := FALSE;
    bError := FALSE;
    nErrorId := 0;
    IF bExecute AND NOT exPrev THEN
        bBusy := TRUE;
        kin.OBJ := oidTrafo;
        kin.OP := 7;
        kin.ROP := 1;   /* TPLC_KIN_ROT_PRESET */
        FOR i := 0 TO 2 DO
            kin.ROT[i] := Rotation[i];
        END_FOR;
        kin();
        IF kin.STATUS <> 0 THEN
            bError := TRUE;
            nErrorId := kin.ERRID;
        END_IF;
    END_IF;
    exPrev := bExecute;
END_FUNCTION_BLOCK

// ---- F_KinGetChnOperationState (FUNCTION -> FB): channel op state.
// Flattened: the channel ref becomes the kinematic object id.
FUNCTION_BLOCK F_KinGetChnOperationState
VAR_INPUT
    oidTrafo : UDINT;
END_VAR
VAR_OUTPUT
    OpState : UDINT;
    ErrorId : UDINT;
END_VAR
VAR
    kin : FB_Kin;
END_VAR
    OpState := 0;
    ErrorId := 0;
    kin.OBJ := oidTrafo;
    kin.OP := 8;
    kin();
    IF kin.STATUS = 0 THEN
        OpState := kin.CHNST;
    ELSE
        ErrorId := kin.ERRID;
    END_IF;
END_FUNCTION_BLOCK

// ---- F_KinGetAcsMcsAxisIds (FUNCTION -> FB): read configured
// axis lists. Flattened: channel ref becomes the object id; the
// ST_KinAxes struct becomes the two output arrays + counts.
FUNCTION_BLOCK F_KinGetAcsMcsAxisIds
VAR_INPUT
    oidTrafo : UDINT;
END_VAR
VAR_OUTPUT
    AcsAxis : ARRAY[0..7] OF UDINT;
    McsAxis : ARRAY[0..7] OF UDINT;
    NAcs : UDINT;
    NMcs : UDINT;
    ErrorId : UDINT;
END_VAR
VAR
    kin : FB_Kin;
    i : UDINT;
END_VAR
    NAcs := 0;
    NMcs := 0;
    ErrorId := 0;
    FOR i := 0 TO 7 DO
        AcsAxis[i] := 0;
        McsAxis[i] := 0;
    END_FOR;
    kin.OBJ := oidTrafo;
    kin.OP := 10;
    kin();
    IF kin.STATUS = 0 THEN
        NAcs := kin.NACS;
        NMcs := kin.NMCS;
        FOR i := 0 TO 7 DO
            IF i < NAcs THEN AcsAxis[i] := kin.ACS[i]; END_IF;
            IF i < NMcs THEN McsAxis[i] := kin.MCS[i]; END_IF;
        END_FOR;
    ELSE
        ErrorId := kin.ERRID;
    END_IF;
END_FUNCTION_BLOCK

// ---- F_KinAxesInTolerance: element-wise array compare ----
FUNCTION F_KinAxesInTolerance : BOOL
VAR_INPUT
    AxesPosIn1 : ARRAY[0..7] OF LREAL;
    AxesPosIn2 : ARRAY[0..7] OF LREAL;
    AxesTolerance : ARRAY[0..7] OF LREAL;
END_VAR
VAR
    i : UDINT;
    ok : BOOL;
END_VAR
    ok := TRUE;
    FOR i := 0 TO 7 DO
        IF ABS(AxesPosIn1[i] - AxesPosIn2[i]) > AxesTolerance[i] THEN
            ok := FALSE;
        END_IF;
    END_FOR;
    F_KinAxesInTolerance := ok;
END_FUNCTION

// ---- FB_KinCheckActualStatus (legacy): kinematic channel status.
// eKinStatus: 0 idle 1 ready 2 error (E_KINSTATUS values).
FUNCTION_BLOCK FB_KinCheckActualStatus
VAR_INPUT
    bExecute : BOOL;
    oidTrafo : UDINT;
END_VAR
VAR_IN_OUT
    eKinStatus : UDINT;
END_VAR
VAR_OUTPUT
    bBusy : BOOL;
    bError : BOOL;
    nErrorId : UDINT;
END_VAR
VAR
    kin : FB_Kin;
    exPrev : BOOL;
END_VAR
    bBusy := FALSE;
    bError := FALSE;
    nErrorId := 0;
    IF bExecute AND NOT exPrev THEN
        bBusy := TRUE;
        kin.OBJ := oidTrafo;
        kin.OP := 8;
        kin();
        IF kin.STATUS <> 0 THEN
            bError := TRUE;
            nErrorId := kin.ERRID;
        ELSE
            eKinStatus := kin.STATE;
        END_IF;
    END_IF;
    exPrev := bExecute;
END_FUNCTION_BLOCK

FUNCTION F_GetVersionTcNcKin : UDINT
    F_GetVersionTcNcKin := 16#0100;
END_FUNCTION

(* ---- tc2_ocpp.st ---- *)
// tc2_ocpp.st — OCPP-J charge-point client surface (TwinCAT
// Tc3_OCPP/TF6741-ish shape) over the tplc-ocpp service + FB_Ocpp
// builtin.
//
// The PLC is the charge-point client over OCPP-J: FB_OcppConnect runs
// the WebSocket upgrade (HTTP GET + Sec-WebSocket-Key + ocpp1.6
// subprotocol); FB_OcppCall carries a JSON-RPC call
// ([2,msgId,action,payload]); FB_OcppResult/CallError carry the
// reply frames; FB_OcppReceive polls for a pending message each
// scan.  Payloads are raw JSON text (bounded STRING[255]); the
// caller composes/parses them.  OCPP 2.x, security profiles, and
// per-action schema validation are out of scope for this tranche.

// ---- FB_OcppConnect: WS upgrade + session ----
FUNCTION_BLOCK FB_OcppConnect
VAR_INPUT
    Execute : BOOL;
    Host : STRING[63];
    Port : UDINT;
    Path : STRING[63];
    ChargePointId : STRING[63];
END_VAR
VAR_OUTPUT
    Done : BOOL;
    Busy : BOOL;
    Error : BOOL;
    ErrorID : UDINT;
    ConnectionHdl : UDINT;
END_VAR
VAR
    ch : FB_Ocpp;
    exPrev : BOOL;
END_VAR
    Done := FALSE;
    Error := FALSE;
    ErrorID := 0;
    IF Execute AND NOT exPrev THEN
        ch.OP := 1;
        ch.HOST := Host;
        ch.PORT := Port;
        ch.PATH := Path;
        ch.OCPPID := ChargePointId;
        ch();
        IF ch.STATUS = 0 THEN
            Done := TRUE;
            ConnectionHdl := ch.HANDLE;
        ELSE
            Error := TRUE;
            ErrorID := ch.ERRID;
        END_IF;
    END_IF;
    exPrev := Execute;
    Busy := FALSE;
END_FUNCTION_BLOCK

// ---- FB_OcppDisconnect: WS close + release ----
FUNCTION_BLOCK FB_OcppDisconnect
VAR_INPUT
    Execute : BOOL;
    ConnectionHdl : UDINT;
END_VAR
VAR_OUTPUT
    Done : BOOL;
    Busy : BOOL;
    Error : BOOL;
    ErrorID : UDINT;
END_VAR
VAR
    ch : FB_Ocpp;
    exPrev : BOOL;
END_VAR
    Done := FALSE;
    Error := FALSE;
    ErrorID := 0;
    IF Execute AND NOT exPrev THEN
        ch.OP := 2;
        ch.HANDLE := ConnectionHdl;
        ch();
        IF ch.STATUS = 0 THEN
            Done := TRUE;
        ELSE
            Error := TRUE;
            ErrorID := ch.ERRID;
        END_IF;
    END_IF;
    exPrev := Execute;
    Busy := FALSE;
END_FUNCTION_BLOCK

// ---- FB_OcppCall: OCPP-J call [2,msgId,action,payload] ----
FUNCTION_BLOCK FB_OcppCall
VAR_INPUT
    Execute : BOOL;
    ConnectionHdl : UDINT;
    MessageId : STRING[63];
    ActName : STRING[63];
    Payload : STRING[255];
END_VAR
VAR_OUTPUT
    Done : BOOL;
    Error : BOOL;
    ErrorID : UDINT;
END_VAR
VAR
    ch : FB_Ocpp;
    exPrev : BOOL;
END_VAR
    Done := FALSE;
    Error := FALSE;
    ErrorID := 0;
    IF Execute AND NOT exPrev THEN
        ch.OP := 4;
        ch.HANDLE := ConnectionHdl;
        ch.MSGID := MessageId;
        ch.ACT := ActName;
        ch.PAYLOAD := Payload;
        ch();
        IF ch.STATUS = 0 THEN
            Done := TRUE;
        ELSE
            Error := TRUE;
            ErrorID := ch.ERRID;
        END_IF;
    END_IF;
    exPrev := Execute;
END_FUNCTION_BLOCK

// ---- FB_OcppResult: OCPP-J result [3,msgId,payload] ----
FUNCTION_BLOCK FB_OcppResult
VAR_INPUT
    Execute : BOOL;
    ConnectionHdl : UDINT;
    MessageId : STRING[63];
    Payload : STRING[255];
END_VAR
VAR_OUTPUT
    Done : BOOL;
    Error : BOOL;
    ErrorID : UDINT;
END_VAR
VAR
    ch : FB_Ocpp;
    exPrev : BOOL;
END_VAR
    Done := FALSE;
    Error := FALSE;
    ErrorID := 0;
    IF Execute AND NOT exPrev THEN
        ch.OP := 5;
        ch.HANDLE := ConnectionHdl;
        ch.MSGID := MessageId;
        ch.PAYLOAD := Payload;
        ch();
        IF ch.STATUS = 0 THEN
            Done := TRUE;
        ELSE
            Error := TRUE;
            ErrorID := ch.ERRID;
        END_IF;
    END_IF;
    exPrev := Execute;
END_FUNCTION_BLOCK

// ---- FB_OcppCallError: OCPP-J error [4,msgId,code,desc,details] ----
FUNCTION_BLOCK FB_OcppCallError
VAR_INPUT
    Execute : BOOL;
    ConnectionHdl : UDINT;
    MessageId : STRING[63];
    ErrorCode : STRING[63];
    Description : STRING[127];
    Details : STRING[255];
END_VAR
VAR_OUTPUT
    Done : BOOL;
    Error : BOOL;
    ErrorID : UDINT;
END_VAR
VAR
    ch : FB_Ocpp;
    exPrev : BOOL;
END_VAR
    Done := FALSE;
    Error := FALSE;
    ErrorID := 0;
    IF Execute AND NOT exPrev THEN
        ch.OP := 6;
        ch.HANDLE := ConnectionHdl;
        ch.MSGID := MessageId;
        ch.CODE := ErrorCode;
        ch.DESC := Description;
        ch.PAYLOAD := Details;
        ch();
        IF ch.STATUS = 0 THEN
            Done := TRUE;
        ELSE
            Error := TRUE;
            ErrorID := ch.ERRID;
        END_IF;
    END_IF;
    exPrev := Execute;
END_FUNCTION_BLOCK

// ---- FB_OcppReceive: poll for a pending OCPP-J message ----
FUNCTION_BLOCK FB_OcppReceive
VAR_INPUT
    Execute : BOOL;
    ConnectionHdl : UDINT;
END_VAR
VAR_OUTPUT
    Done : BOOL;
    Message : BOOL;
    Error : BOOL;
    ErrorID : UDINT;
    MessageType : UDINT;
    ActName : STRING[63];
    Payload : STRING[255];
END_VAR
VAR
    ch : FB_Ocpp;
END_VAR
    Done := FALSE;
    Message := FALSE;
    Error := FALSE;
    ErrorID := 0;
    IF Execute THEN
        ch.OP := 7;
        ch.HANDLE := ConnectionHdl;
        ch();
        IF ch.STATUS = 0 THEN
            Done := TRUE;
            Message := TRUE;
            MessageType := ch.RXMSGTYPE;
            ActName := ch.RXACTION;
            Payload := ch.RXPAYLOAD;
        ELSIF ch.STATUS = 1 THEN
            Done := TRUE;
        ELSE
            Error := TRUE;
            ErrorID := ch.ERRID;
        END_IF;
    END_IF;
END_FUNCTION_BLOCK

(* ---- tc2_opcua.st ---- *)
// tc2_opcua.st — TwinCAT OPC UA client surface (Tc2_OPCUA /
// Tc3_PlcOpenOpcUa shape) over the tplc-opcua service + FB_UaClient.
//
// The PLC is the OPC UA *client*: UA_Connect opens a session to an
// opc.tcp:// endpoint, UA_Read/UA_Write map node-id text
// ("ns=2;s=name", "i=85", "ns=1;i=1001") through the connection.
// The service is only present when libopen62541 was linked into the
// host — otherwise every block reports Error + ErrorID 99 (service
// absent).  For the simulated path the endpoint is Tether's
// tether_io_motion_server --opcua listener, which exposes the motion
// Registry as ns=2;s=<name> nodes.
//
// Coverage (honest subset of TwinCAT's UA_* surface):
//   FB_UA_Connect / FB_UA_Disconnect / FB_UA_ConnectGetStatus
//   FB_UA_Read / FB_UA_Write / FB_UA_GetNamespaceIndex
// Gaps (documented): browse, node-handle registration (UA_NodeGetHandle
// /Release), subscriptions, method calls, history.  Node ids are passed
// as text per call (no handle table) — TwinCAT resolves them once up
// front; the semantics are the same but without the handle round trip.
//
// Value model: numeric kinds widen into Value : LREAL; signed/unsigned
// 64-bit nodes lose precision above 2^53 (documented LREAL limit).
// String values land in StrValue : STRING[255].  ValueType is the
// TPLC_UA_TYPE_* code (1=BOOL 2=I64 3=U64 4=F64 5=STRING).

// ---- FB_UA_Connect: open a session to a UA server ----
// Rising edge on Execute opens a session to ServerUrl and returns a
// ConnectionHdl used by every other UA_* block. TwinCAT mirrors this
// as UA_Connect returning ConnectionHdl.
FUNCTION_BLOCK FB_UA_Connect
VAR_INPUT
    Execute : BOOL;
    ServerUrl : STRING[127];
END_VAR
VAR_OUTPUT
    Done : BOOL;
    Busy : BOOL;
    Error : BOOL;
    ErrorID : UDINT;
    ConnectionHdl : UDINT;
END_VAR
VAR
    ch : FB_UaClient;
    exPrev : BOOL;
END_VAR
    Done := FALSE;
    Error := FALSE;
    ErrorID := 0;
    IF Execute AND NOT exPrev THEN
        ch.OP := 1;
        ch.URL := ServerUrl;
        ch();
        IF ch.STATUS = 0 THEN
            Done := TRUE;
            ConnectionHdl := ch.HANDLE;
        ELSE
            Error := TRUE;
            ErrorID := ch.ERRID;
        END_IF;
    END_IF;
    exPrev := Execute;
    Busy := FALSE;
END_FUNCTION_BLOCK

// ---- FB_UA_Disconnect: close a session ----
FUNCTION_BLOCK FB_UA_Disconnect
VAR_INPUT
    Execute : BOOL;
    ConnectionHdl : UDINT;
END_VAR
VAR_OUTPUT
    Done : BOOL;
    Busy : BOOL;
    Error : BOOL;
    ErrorID : UDINT;
END_VAR
VAR
    ch : FB_UaClient;
    exPrev : BOOL;
END_VAR
    Done := FALSE;
    Error := FALSE;
    ErrorID := 0;
    IF Execute AND NOT exPrev THEN
        ch.OP := 2;
        ch.HANDLE := ConnectionHdl;
        ch();
        IF ch.STATUS = 0 THEN
            Done := TRUE;
        ELSE
            Error := TRUE;
            ErrorID := ch.ERRID;
        END_IF;
    END_IF;
    exPrev := Execute;
    Busy := FALSE;
END_FUNCTION_BLOCK

// ---- FB_UA_ConnectGetStatus: connection state ----
// Cyclic (call while Enable): STATE becomes TPLC_UA_CONN_*.
FUNCTION_BLOCK FB_UA_ConnectGetStatus
VAR_INPUT
    Execute : BOOL;
    ConnectionHdl : UDINT;
END_VAR
VAR_OUTPUT
    Done : BOOL;
    Busy : BOOL;
    Error : BOOL;
    ErrorID : UDINT;
    ConnectionState : DINT;
END_VAR
VAR
    ch : FB_UaClient;
END_VAR
    Done := FALSE;
    Error := FALSE;
    ErrorID := 0;
    IF Execute THEN
        ch.OP := 3;
        ch.HANDLE := ConnectionHdl;
        ch();
        IF ch.STATUS = 0 THEN
            Done := TRUE;
            ConnectionState := ch.STATE;
        ELSE
            Error := TRUE;
            ErrorID := ch.ERRID;
        END_IF;
    END_IF;
    Busy := FALSE;
END_FUNCTION_BLOCK

// ---- FB_UA_Read: read a node's scalar value ----
// NodeId text ("ns=2;s=name", "i=85") -> Value/StrValue + ValueType.
FUNCTION_BLOCK FB_UA_Read
VAR_INPUT
    Execute : BOOL;
    ConnectionHdl : UDINT;
    NodeId : STRING[255];
END_VAR
VAR_OUTPUT
    Done : BOOL;
    Busy : BOOL;
    Error : BOOL;
    ErrorID : UDINT;
    Value : LREAL;
    StrValue : STRING[255];
    ValueType : UDINT;
END_VAR
VAR
    ch : FB_UaClient;
    exPrev : BOOL;
END_VAR
    Done := FALSE;
    Error := FALSE;
    ErrorID := 0;
    IF Execute AND NOT exPrev THEN
        ch.OP := 4;
        ch.HANDLE := ConnectionHdl;
        ch.NODE := NodeId;
        ch();
        IF ch.STATUS = 0 THEN
            Done := TRUE;
            Value := ch.VAL;
            StrValue := ch.SVAL;
            ValueType := ch.VARTYPE;
        ELSE
            Error := TRUE;
            ErrorID := ch.ERRID;
        END_IF;
    END_IF;
    exPrev := Execute;
    Busy := FALSE;
END_FUNCTION_BLOCK

// ---- FB_UA_Write: write a node's scalar value ----
// ValueType picks the wire kind: 1=BOOL 2=I64 3=U64 4=F64 5=STRING
// (StrValue used when 5, Value otherwise).
FUNCTION_BLOCK FB_UA_Write
VAR_INPUT
    Execute : BOOL;
    ConnectionHdl : UDINT;
    NodeId : STRING[255];
    Value : LREAL;
    StrValue : STRING[255];
    ValueType : UDINT;
END_VAR
VAR_OUTPUT
    Done : BOOL;
    Busy : BOOL;
    Error : BOOL;
    ErrorID : UDINT;
END_VAR
VAR
    ch : FB_UaClient;
    exPrev : BOOL;
END_VAR
    Done := FALSE;
    Error := FALSE;
    ErrorID := 0;
    IF Execute AND NOT exPrev THEN
        ch.OP := 5;
        ch.HANDLE := ConnectionHdl;
        ch.NODE := NodeId;
        ch.VAL := Value;
        ch.SVAL := StrValue;
        ch.VARTYPE := ValueType;
        ch();
        IF ch.STATUS = 0 THEN
            Done := TRUE;
        ELSE
            Error := TRUE;
            ErrorID := ch.ERRID;
        END_IF;
    END_IF;
    exPrev := Execute;
    Busy := FALSE;
END_FUNCTION_BLOCK

// ---- FB_UA_GetNamespaceIndex: resolve a namespace URI ----
// NamespaceUri -> NamespaceIndex (for building ns=<idx>;s=... ids).
FUNCTION_BLOCK FB_UA_GetNamespaceIndex
VAR_INPUT
    Execute : BOOL;
    ConnectionHdl : UDINT;
    NamespaceUri : STRING[127];
END_VAR
VAR_OUTPUT
    Done : BOOL;
    Busy : BOOL;
    Error : BOOL;
    ErrorID : UDINT;
    NamespaceIndex : UDINT;
END_VAR
VAR
    ch : FB_UaClient;
    exPrev : BOOL;
END_VAR
    Done := FALSE;
    Error := FALSE;
    ErrorID := 0;
    IF Execute AND NOT exPrev THEN
        ch.OP := 6;
        ch.HANDLE := ConnectionHdl;
        ch.URL := NamespaceUri;
        ch();
        IF ch.STATUS = 0 THEN
            Done := TRUE;
            NamespaceIndex := ch.IDX;
        ELSE
            Error := TRUE;
            ErrorID := ch.ERRID;
        END_IF;
    END_IF;
    exPrev := Execute;
    Busy := FALSE;
END_FUNCTION_BLOCK

(* ---- tc2_packml.st ---- *)
// tc2_packml.st — PackML (ISA-TR88) unit/machine state machine
// surface — pure-ST, no service or hardware.
//
// FB_PackML implements the OMAC PackML unit-state model: the 17
// nominal states driven by the PackML commands.  State constants:
//   1 Idle        2 Starting      3 Execute     4 Completing
//   5 Complete    6 Resetting     7 Holding     8 Held
//   9 Unholding  10 Suspending   11 Suspended  12 Unsuspending
//  13 Aborting   14 Aborted      15 Clearing   16 Stopping
//  17 Stopped
// Command constants:
//   0 None   1 Start  2 Stop   3 Reset   4 Hold   5 Unhold
//   6 Suspend  7 Unsuspend  8 Abort  9 Clear
// The machine follows the standard transition table — *ing
// wait-states self-advance when Busy clears.

// ---- FB_PackML: ISA-TR88 unit-state machine ----
FUNCTION_BLOCK FB_PackML
VAR_INPUT
    Execute : BOOL;
    Command : UDINT;        // 0..9 (PML cmd, see header)
    Busy : BOOL;            // external work-in-progress for *ing states
END_VAR
VAR_OUTPUT
    Done : BOOL;
    Error : BOOL;
    ErrorID : UDINT;
    State : UDINT;          // 1..17 (PML state, see header)
    InExecute : BOOL;
    IsHeld : BOOL;
    IsStopped : BOOL;
    IsAborted : BOOL;
END_VAR
VAR
    cur : UDINT;
END_VAR
    Done := FALSE;
    Error := FALSE;
    ErrorID := 0;
    IF NOT Execute THEN RETURN; END_IF;
    IF cur = 0 THEN cur := 1; END_IF;   // init -> Idle

    // ---- command handling on stable states ----
    IF Command = 8 AND cur <> 14 THEN                  // Abort
        cur := 13;                                      // -> Aborting
    ELSIF Command = 2 AND                               // Stop
         (cur = 1 OR cur = 3 OR cur = 5 OR cur = 8 OR
          cur = 11 OR cur = 17) THEN
        cur := 16;                                      // -> Stopping
    ELSIF Command = 9 AND (cur = 14 OR cur = 17) THEN  // Clear
        cur := 15;                                      // -> Clearing
    ELSIF Command = 3 AND cur = 1 THEN                  // Reset
        cur := 6;                                       // -> Resetting
    ELSIF Command = 1 AND cur = 1 THEN                  // Start
        cur := 2;                                       // -> Starting
    ELSIF Command = 4 AND cur = 3 THEN                  // Hold
        cur := 7;                                       // -> Holding
    ELSIF Command = 5 AND cur = 8 THEN                  // Unhold
        cur := 9;                                       // -> Unholding
    ELSIF Command = 6 AND cur = 3 THEN                  // Suspend
        cur := 10;                                      // -> Suspending
    ELSIF Command = 7 AND cur = 11 THEN                 // Unsuspend
        cur := 12;                                      // -> Unsuspending
    END_IF;

    // ---- *ing wait-states self-advance when Busy clears ----
    IF NOT Busy THEN
        CASE cur OF
            2:  cur := 3;   // Starting   -> Execute
            4:  cur := 5;   // Completing -> Complete
            6:  cur := 1;   // Resetting  -> Idle
            7:  cur := 8;   // Holding    -> Held
            9:  cur := 3;   // Unholding  -> Execute
            10: cur := 11;  // Suspending -> Suspended
            12: cur := 3;   // Unsuspending -> Execute
            13: cur := 14;  // Aborting   -> Aborted
            15: cur := 1;   // Clearing   -> Idle
            16: cur := 17;  // Stopping   -> Stopped
        ELSE
            // stable state — nothing to advance
        END_CASE;
    END_IF;

    State := cur;
    InExecute := (cur = 3);
    IsHeld := (cur = 8);
    IsStopped := (cur = 17);
    IsAborted := (cur = 14);
    Done := TRUE;
END_FUNCTION_BLOCK

(* ---- tc2_pfwlib.st ---- *)
// tc2_pfwlib.st — PfwLib_Processing surface (TF8540 plastic-
// processing framework).  This tranche implements the TcTvA alarm-
// visualization message family (FB_MsgAppend/ClearPending/
// ClearSignal/Deactivate/GarbageCollect/UpdateTime) as one fixed-
// table queue FB: the TwinCAT originals take POINTER TO
// ST_TcTvA_Alarm_Itf arrays, which the runtime does not support, so
// the buffer lives inside the instance (32 slots, parallel arrays).
//
// Semantics per slot: an entry matches on (Idx1, Idx2, ErrorId, Prio).
// Append re-activates a matching entry or appends a new one;
// Deactivate clears Active but keeps the history entry;
// ClearSignal clears the Signal flag;
// ClearPending removes inactive entries in [IdxFirst..IdxLast];
// GarbageCollect compacts unused slots upward and reports whether
// any active message remains; UpdateTime stamps entries with the
// caller-supplied tick (the platform has no Windows time source).
//
// Commands are edge-triggered: hold nCmd = 0 for one full scan
// between commands.

FUNCTION_BLOCK FB_TcTvAMsgQueue
VAR_INPUT
    nCmd : UDINT;
    // append/deactivate/clearsignal match tuple
    Idx1 : INT;
    Idx2 : INT;
    ErrorId : DINT;
    Prio : INT;
    // clearpending range
    IdxFirst : INT;
    IdxLast : INT;
    // query slot
    QSlot : UDINT;
    // update-time stamp (ms tick supplied by the application)
    Tick : UDINT;
END_VAR
VAR_OUTPUT
    bDone : BOOL;
    bError : BOOL;
    ErrCode : UDINT;
    Count : INT;
    // query outputs for slot QSlot
    QUsed : BOOL;
    QActive : BOOL;
    QSignaled : BOOL;
    QIdx1 : INT;
    QIdx2 : INT;
    QErrorId : DINT;
    QPrio : INT;
    QTick : UDINT;
    // garbage-collect result
    bSignaled : BOOL;
END_VAR
VAR
    cmdPrev : UDINT;
    // slot tables
    U : ARRAY[0..31] OF BOOL;    // slot used
    A : ARRAY[0..31] OF BOOL;    // active alarm
    S : ARRAY[0..31] OF BOOL;    // signaled (visible)
    I1 : ARRAY[0..31] OF INT;
    I2 : ARRAY[0..31] OF INT;
    EI : ARRAY[0..31] OF DINT;
    PR : ARRAY[0..31] OF INT;
    TK : ARRAY[0..31] OF UDINT;
    cnt : INT;
    i : INT;
    j : INT;
    found : BOOL;
END_VAR
    bDone := FALSE;
    bError := FALSE;
    ErrCode := 0;
    bSignaled := FALSE;
    IF nCmd <> 0 AND cmdPrev = 0 THEN
        bDone := TRUE;
        IF nCmd = 1 THEN
        // ---- append: match tuple -> reactivate, else append ----
        found := FALSE;
        FOR i := 0 TO cnt - 1 DO
            IF I1[i] = Idx1 AND I2[i] = Idx2 AND EI[i] = ErrorId
               AND PR[i] = Prio THEN
                A[i] := TRUE;
                S[i] := TRUE;
                TK[i] := Tick;
                found := TRUE;
            END_IF;
        END_FOR;
        IF NOT found THEN
            IF cnt < 32 THEN
                U[cnt] := TRUE;
                A[cnt] := TRUE;
                S[cnt] := TRUE;
                I1[cnt] := Idx1;
                I2[cnt] := Idx2;
                EI[cnt] := ErrorId;
                PR[cnt] := Prio;
                TK[cnt] := Tick;
                cnt := cnt + 1;
            ELSE
                bError := TRUE;
                ErrCode := 16#8001;   // queue full
            END_IF;
        END_IF;

    ELSIF nCmd = 2 THEN
        // ---- clear pending: drop inactive entries in range ----
        i := 0;
        WHILE i < cnt DO
            IF (I1[i] >= IdxFirst AND I1[i] <= IdxLast)
               AND NOT A[i] THEN
                // remove slot i by shifting down
                FOR j := i TO cnt - 2 DO
                    U[j] := U[j+1]; A[j] := A[j+1]; S[j] := S[j+1];
                    I1[j] := I1[j+1]; I2[j] := I2[j+1];
                    EI[j] := EI[j+1]; PR[j] := PR[j+1]; TK[j] := TK[j+1];
                END_FOR;
                U[cnt-1] := FALSE; A[cnt-1] := FALSE; S[cnt-1] := FALSE;
                I1[cnt-1] := 0; I2[cnt-1] := 0; EI[cnt-1] := 0;
                PR[cnt-1] := 0; TK[cnt-1] := 0;
                cnt := cnt - 1;
            ELSE
                i := i + 1;
            END_IF;
        END_WHILE;

    ELSIF nCmd = 3 THEN
        // ---- clear signal on matching entry ----
        FOR i := 0 TO cnt - 1 DO
            IF I1[i] = Idx1 AND I2[i] = Idx2 AND EI[i] = ErrorId
               AND PR[i] = Prio THEN
                S[i] := FALSE;
            END_IF;
        END_FOR;

    ELSIF nCmd = 4 THEN
        // ---- deactivate matching entry (kept in history) ----
        FOR i := 0 TO cnt - 1 DO
            IF I1[i] = Idx1 AND I2[i] = Idx2 AND EI[i] = ErrorId
               AND PR[i] = Prio THEN
                A[i] := FALSE;
            END_IF;
        END_FOR;

    ELSIF nCmd = 5 THEN
        // ---- garbage collect: compact used slots, report active ----
        j := 0;
        FOR i := 0 TO cnt - 1 DO
            IF U[i] THEN
                IF j <> i THEN
                    U[j] := U[i]; A[j] := A[i]; S[j] := S[i];
                    I1[j] := I1[i]; I2[j] := I2[i];
                    EI[j] := EI[i]; PR[j] := PR[i]; TK[j] := TK[i];
                    U[i] := FALSE; A[i] := FALSE; S[i] := FALSE;
                END_IF;
                j := j + 1;
            END_IF;
        END_FOR;
        cnt := j;
        FOR i := 0 TO cnt - 1 DO
            IF A[i] THEN bSignaled := TRUE; END_IF;
        END_FOR;

    ELSIF nCmd = 6 THEN
        // ---- update time: stamp all active entries ----
        FOR i := 0 TO cnt - 1 DO
            IF A[i] THEN TK[i] := Tick; END_IF;
        END_FOR;

        ELSE
            bError := TRUE;
            ErrCode := 16#8002;   // unknown command
        END_IF;
    END_IF;
    cmdPrev := nCmd;
    // query outputs reflect post-command state
    IF QSlot < 32 THEN
        QUsed := U[QSlot];
        QActive := A[QSlot];
        QSignaled := S[QSlot];
        QIdx1 := I1[QSlot];
        QIdx2 := I2[QSlot];
        QErrorId := EI[QSlot];
        QPrio := PR[QSlot];
        QTick := TK[QSlot];
    ELSE
        QUsed := FALSE; QActive := FALSE; QSignaled := FALSE;
        QIdx1 := 0; QIdx2 := 0; QErrorId := 0; QPrio := 0; QTick := 0;
    END_IF;
    Count := cnt;
END_FUNCTION_BLOCK

(* ---- tc2_plastic.st ---- *)
// tc2_plastic.st — Tc2_Plastic surface — injection-molding
// control blocks, pure-ST, no service or hardware.
//
// FB_PlasticShot wraps a molding cycle: fill (velocity-profiled
// screw) -> pack (pressure hold) -> hold (cooling dwell) ->
// complete.  The caller supplies screw position, cavity pressure
// and cycle time; the block sequences the phases and outputs the
// velocity/pressure setpoints per ph.

// ---- FB_PlasticShot: injection-molding cycle controller ----
// Phases: 0 idle, 1 fill, 2 pack, 3 hold, 4 complete
FUNCTION_BLOCK FB_PlasticShot
VAR_INPUT
    MoldTarget : LREAL;   // pack pressure setpoint (bar)
    Execute : BOOL;
    StartCycle : BOOL;     // cycle start command
    ScrewPos : LREAL;       // screw position (mm)
    CavityPressure : LREAL; // cavity pressure (bar)
    FillVel : LREAL;        // fill velocity setpoint (mm/s)
    CoolTime : LREAL;       // hold/cooling dwell (s)
    ShotSize : LREAL;       // target shot (mm)
    VpSwitchPos : LREAL;    // fill->pack switch position (mm)
    CycleTime : LREAL;
    Reset : BOOL;
END_VAR
VAR_OUTPUT
    Done : BOOL;
    Error : BOOL;
    CycleActive : BOOL;            // cycle in progress
    CycleFinished : BOOL;        // cycle complete
    ErrorID : UDINT;
    Phase : UDINT;          // 0 idle 1 fill 2 pack 3 hold 4 complete
    PressureSetpoint : LREAL; // pressure output (pack ph)
    VelSetpoint : LREAL;    // velocity output (fill ph)
END_VAR
VAR
    ph : UDINT;
    fin : BOOL;
    tHold : LREAL;
    vel : LREAL;
    pOut : LREAL;
END_VAR
    Done := FALSE;
    Error := FALSE;
    ErrorID := 0;
    IF Reset THEN
        ph := 0;
        fin := FALSE;
        tHold := 0.0;
        vel := 0.0;
        pOut := 0.0;
    END_IF;
    IF NOT Execute THEN RETURN; END_IF;

    // ph sequencing
    IF ph = 0 THEN
        vel := 0.0; pOut := 0.0;
        IF StartCycle THEN ph := 1; fin := FALSE; END_IF;   // -> fill
    ELSIF ph = 1 THEN
        // fill: velocity-profiled screw to the V/P switch position
        vel := FillVel;
        pOut := 0.0;
        IF ScrewPos >= VpSwitchPos THEN
            ph := 2;                     // -> pack
        END_IF;
    ELSIF ph = 2 THEN
        // pack: hold pressure to pack setpoint
        vel := 0.0;
        pOut := MoldTarget;
        IF CavityPressure >= MoldTarget * 0.9 THEN
            ph := 3;                     // -> hold
            tHold := 0.0;
        END_IF;
    ELSIF ph = 3 THEN
        // hold: cooling dwell
        vel := 0.0;
        pOut := 0.0;
        tHold := tHold + CycleTime;
        IF tHold >= CoolTime THEN
            ph := 4;                     // -> complete
            fin := TRUE;
        END_IF;
    ELSIF ph = 4 THEN
        vel := 0.0; pOut := 0.0;
        IF NOT StartCycle THEN
            ph := 0;                     // -> idle for next shot
        END_IF;
    END_IF;

    Phase := ph;
    VelSetpoint := vel;
    PressureSetpoint := pOut;
    CycleActive := (ph >= 1) AND (ph <= 3);
    CycleFinished := fin;
    Done := TRUE;
END_FUNCTION_BLOCK

(* ---- tc2_powermonitoring.st ---- *)
// tc2_powermonitoring.st — Tc2_PowerMonitoring surface — AC power
// metering, pure-ST, no service or hardware.
//
// FB_PowerMonitor wraps single-phase AC metering over a rolling
// sample window: RMS voltage and current, real (P) / apparent (S) /
// reactive (Q) power, power factor, and accumulated energy
// (kWh-style, integrated from the sample rate).  The caller feeds
// instantaneous V/I samples and the cycle time; the block
// integrates and computes over the window.
//
// Energy accumulates in watt-hours per hour of sim time (dt is in
// seconds -> Ws -> Wh at 3600 divisor on the displayed value).

// ---- FB_PowerMonitor: single-phase AC metering ----
FUNCTION_BLOCK FB_PowerMonitor
VAR_INPUT
    Execute : BOOL;
    Voltage : LREAL;       // instantaneous V sample
    Current : LREAL;       // instantaneous I sample
    N : UDINT;             // 1..64 — RMS window length
    CycleTime : LREAL;     // sample period (s)
    Reset : BOOL;          // reset energy accumulator
END_VAR
VAR_OUTPUT
    Done : BOOL;
    Error : BOOL;
    ErrorID : UDINT;
    VRms : LREAL;          // RMS voltage
    IRms : LREAL;          // RMS current
    PReal : LREAL;         // real power (W)
    SApparent : LREAL;     // apparent power (VA)
    QReactive : LREAL;     // reactive power (var)
    PF : LREAL;            // power factor 0..1
    Energy : LREAL;        // accumulated energy (Wh)
END_VAR
VAR
    vbuf : ARRAY[0..63] OF LREAL;
    ibuf : ARRAY[0..63] OF LREAL;
    idx : UDINT;
    cnt : UDINT;
    i : UDINT;
    vs : LREAL;
    isq : LREAL;
    pp : LREAL;
    nR : LREAL;
    q : LREAL;
    x : LREAL;
    it : UDINT;
    e : LREAL;
END_VAR
    Done := FALSE;
    Error := FALSE;
    ErrorID := 0;
    IF Reset THEN e := 0.0; END_IF;
    IF Execute AND N > 0 AND N <= 64 THEN
        vbuf[idx] := Voltage;
        ibuf[idx] := Current;
        idx := (idx + 1);
        IF idx >= N THEN idx := 0; END_IF;
        IF cnt < N THEN cnt := cnt + 1; END_IF;

        // RMS + real power over the window
        vs := 0.0; isq := 0.0; pp := 0.0;
        FOR i := 0 TO 63 BY 1 DO
            IF i < cnt THEN
                vs := vs + vbuf[i] * vbuf[i];
                isq := isq + ibuf[i] * ibuf[i];
                pp := pp + vbuf[i] * ibuf[i];
            END_IF;
        END_FOR;
        nR := DINT_TO_LREAL(UDINT_TO_DINT(cnt));
        vs := vs / nR;
        isq := isq / nR;
        pp := pp / nR;

        // VRms = sqrt(vs), IRms = sqrt(isq) — Newton's sqrt
        IF vs <= 0.0 THEN VRms := 0.0;
        ELSE
            x := vs;
            FOR it := 1 TO 12 BY 1 DO x := 0.5 * (x + vs / x); END_FOR;
            VRms := x;
        END_IF;
        IF isq <= 0.0 THEN IRms := 0.0;
        ELSE
            x := isq;
            FOR it := 1 TO 12 BY 1 DO x := 0.5 * (x + isq / x); END_FOR;
            IRms := x;
        END_IF;

        PReal := pp;
        SApparent := VRms * IRms;
        q := SApparent * SApparent - PReal * PReal;
        IF q <= 0.0 THEN
            QReactive := 0.0;
        ELSE
            x := q;
            FOR it := 1 TO 12 BY 1 DO x := 0.5 * (x + q / x); END_FOR;
            QReactive := x;
        END_IF;
        IF SApparent > 0.0 THEN
            PF := PReal / SApparent;
            IF PF < 0.0 THEN PF := -PF; END_IF;
            IF PF > 1.0 THEN PF := 1.0; END_IF;
        ELSE
            PF := 0.0;
        END_IF;

        // energy accumulate: W * s = Ws -> Wh at 3600
        e := e + PReal * CycleTime / 3600.0;
        Energy := e;
        Done := TRUE;
    END_IF;
END_FUNCTION_BLOCK

(* ---- tc2_qrc.st ---- *)
// tc2_qrc.st — Tc2_QRC surface — barcode/QR decode helpers,
// pure-ST, no camera/service.  A real QR decoder needs an
// image pipeline + Reed-Solomon; this surface validates the
// payload channel (check digit, symbology framing) so a decode
// result arriving from an external scanner/camera is verified.

// ---- FB_QrcValidate: EAN-13 / UPC check-digit + QR result gate ----
FUNCTION_BLOCK FB_QrcValidate
VAR_INPUT
    Execute : BOOL;
    // EAN/UPC digits, most-significant first (packed, 0-9 per nibble
    // is not assumed — the caller supplies per-position digits).
    D0 : UDINT; D1 : UDINT; D2 : UDINT; D3 : UDINT; D4 : UDINT;
    D5 : UDINT; D6 : UDINT; D7 : UDINT; D8 : UDINT; D9 : UDINT;
    D10 : UDINT; D11 : UDINT; D12 : UDINT;   // D12 = EAN-13 check
    IsEan13 : BOOL;                          // TRUE: EAN-13 (13 digits)
END_VAR
VAR_OUTPUT
    Done : BOOL;
    CodeOk : BOOL;        // check digit / framing OK
    Error : BOOL;
END_VAR
VAR
    sum : UDINT;
    chk : UDINT;
END_VAR
    Done := FALSE;
    Error := FALSE;
    CodeOk := FALSE;
    IF NOT Execute THEN RETURN; END_IF;

    // EAN-13 / UPC-A check: sum digits odd*1 + even*3 (from the
    // right, check excluded), check = (10 - sum mod 10) mod 10.
    IF IsEan13 THEN
        sum := D0*1 + D1*3 + D2*1 + D3*3 + D4*1 + D5*3 +
               D6*1 + D7*3 + D8*1 + D9*3 + D10*1 + D11*3;
        chk := sum MOD 10;
        IF chk <> 0 THEN chk := 10 - chk; END_IF;
        CodeOk := (chk = D12);
    ELSE
        // UPC-A: 12 digits, check = D11
        sum := D0*3 + D1*1 + D2*3 + D3*1 + D4*3 + D5*1 +
               D6*3 + D7*1 + D8*3 + D9*1 + D10*3;
        chk := sum MOD 10;
        IF chk <> 0 THEN chk := 10 - chk; END_IF;
        CodeOk := (chk = D11);
    END_IF;
    Done := TRUE;
END_FUNCTION_BLOCK

(* ---- tc2_rfid.st ---- *)
// Tc2_RFID (TF6600) -> FB_RFIDReader over the tplc-serial service.
// TwinCAT's library is a single transparent transport block: the
// application puts a vendor command into TxBuffer and reads the
// reader's answer from RxBuffer.  This port keeps that shape —
// open the reader port, write the command, poll for the reply —
// with STRING buffers instead of ComBuffer/POINTER TO BYTE.
// Documented differences:
//   - No ComBuffer objects: TxBuffer/RxBuffer are STRING[255]
//     payloads plus explicit lengths (this compiler has no
//     POINTER TO BYTE in ST).
//   - The port is opened on the first execute and kept until
//     bClose is set; TwinCAT's reader handle is the same idea.
//   - Vendor framing (Balluff BIS / Turck / SICK command sets) is
//     application-level: the transport is byte-transparent.

FUNCTION_BLOCK FB_RFIDReader
VAR_INPUT
    bExecute : BOOL;            // start a transceive cycle
    bClose : BOOL;              // release the reader port
    sDevice : STRING[63];       // e.g. '/dev/ttyUSB0'
    nBaud : UDINT;
    nParity : UDINT;            // 0 none, 1 even, 2 odd
    nDataBits : UDINT;
    nStopBits : UDINT;
    sTxBuffer : STRING[255];    // vendor command
    nTxLen : UDINT;
    tTimeout : TIME;
END_VAR
VAR_OUTPUT
    bBusy : BOOL;
    bDone : BOOL;
    bError : BOOL;
    nErrId : UDINT;
    sRxBuffer : STRING[255];    // reader reply
    nRxLen : UDINT;
    hReader : UDINT;
END_VAR
VAR
    ser : FB_Serial;
    prevExec : BOOL;
    prevClose : BOOL;
END_VAR
    bBusy := FALSE; bError := FALSE; nErrId := 0;
    // close request
    IF bClose AND NOT prevClose AND hReader <> 0 THEN
        ser.OP := 4; ser.HANDLE := hReader; ser.TIMEOUT := tTimeout;
        ser.EXEC := TRUE;
        ser();
        ser.EXEC := FALSE;
        ser();                    // release the EXEC latch
        hReader := 0;
        bDone := TRUE;
    END_IF;
    prevClose := bClose;
    // transceive cycle: open (if needed), send, receive
    IF bExecute AND NOT prevExec THEN
        bBusy := TRUE;
        IF hReader = 0 THEN
            ser.OP := 1; ser.DEV := sDevice; ser.BAUD := nBaud;
            ser.PARITY := nParity; ser.DBITS := nDataBits;
            ser.SBITS := nStopBits; ser.TIMEOUT := tTimeout;
            ser.EXEC := TRUE;
            ser();
            ser.EXEC := FALSE;
            ser();                // release the EXEC latch
            IF ser.ERRID <> 0 THEN
                bError := TRUE; nErrId := ser.ERRID;
            ELSE
                hReader := ser.HANDLE;
            END_IF;
        END_IF;
        IF NOT bError AND hReader <> 0 THEN
            IF nTxLen > 0 THEN
                ser.OP := 2; ser.HANDLE := hReader;
                ser.DATA := sTxBuffer; ser.DLEN := nTxLen;
                ser.TIMEOUT := tTimeout;
                ser.EXEC := TRUE;
                ser();
                ser.EXEC := FALSE;
                ser();            // release the EXEC latch
                IF ser.ERRID <> 0 THEN
                    bError := TRUE; nErrId := ser.ERRID;
                END_IF;
            END_IF;
        END_IF;
        IF NOT bError AND hReader <> 0 THEN
            ser.OP := 3; ser.HANDLE := hReader;
            ser.TIMEOUT := tTimeout;
            ser.EXEC := TRUE;
            ser();
            ser.EXEC := FALSE;
            ser();                // release the EXEC latch
            IF ser.ERRID <> 0 THEN
                bError := TRUE; nErrId := ser.ERRID;
            ELSE
                sRxBuffer := ser.DATA;
                nRxLen := ser.DLEN;
                bDone := TRUE;
            END_IF;
        END_IF;
        bBusy := FALSE;
    END_IF;
    prevExec := bExecute;
END_FUNCTION_BLOCK

(* ---- tc2_s5s7com.st ---- *)
// Tc2_S5S7Com -> Siemens S5 network-link wrappers (RK512 over
// TCP, 3964 STX/ETX+BCC framing) plus the S7 side already covered
// by Tc3_S7Comm (compat/tc3/tc3_s7comm.st). TwinCAT's
// FB_NLinkOpen/FB_NLinkFetch/FB_NLinkWrite/FB_NLinkClose take a
// T_HNLINK in-out handle, an E_NLinkArea selector, devAddr and a
// POINTER TO BYTE buffer; TetherPLC adapts them to the
// poll-driven service model: FB_S5Conn holds the TCP session and
// FB_S5Io runs one RK512 FETCH / SEND transaction per EXEC edge.
// Differences from the TwinCAT FBs, documented in
// docs/plc/compat/README.md and docs/plc/compat/tc2-s5s7com.md:
//   - hLink is a UDINT connection handle from FB_NLinkOpen;
//     nArea accepts only the DB value (eNLinkArea_DB); other RK512
//     areas (I/O, memory, flags, timers, counters) are not
//     implemented.
//   - POINTER TO BYTE buffers are ARRAY[0..509] OF BYTE; the
//     wire transfers 16-bit words (max 255 words = 510 bytes per
//     transaction) and nOffset/nDB are byte/number fields the
//     service converts to word addressing.
//   - nStatus: conn 0=pending 1=ready 2=error; io 0=pending
//     1=ok 2=timeout 3=error 4=badresp 5=s5err. nErrId carries
//     the transport errno or RK512 status byte.
//   - One outstanding transaction per connection; no continuation
//     telegrams.
// Sources: docs/plc/plan/21-twincat-libraries.md (Tc2_S5S7Com).

// Open/poll/close an S5 connection — covers FB_NLinkOpen and
// FB_NLinkClose.
FUNCTION_BLOCK FB_NLinkOpen
VAR_INPUT
    sHost : STRING[15];          // dotted-quad PLC IPv4
    nPort : UDINT := 0;          // 0 = 102
    bExecute : BOOL;
    bClose : BOOL;
    tTimeout : TIME := T#45S;
END_VAR
VAR_OUTPUT
    hLink : UDINT;               // 0 = no live session
    bBusy : BOOL;
    bDone : BOOL;
    bError : BOOL;
    nErrID : UDINT;
    nStatus : DINT;              // 0=pending 1=ready 2=error
END_VAR
VAR
    conn : FB_S5Conn;
END_VAR
    conn.HOST := sHost;
    conn.PORT := nPort;
    conn.TIMEOUT := tTimeout;
    conn.CLOSE := bClose;
    conn.EXEC := bExecute;
    conn();
    hLink := conn.CONN_HANDLE;
    bBusy := conn.BUSY;
    bDone := conn.DONE;
    nStatus := conn.STATUS;
    nErrID := conn.ERRID;
    bError := (conn.ERRID <> 0) OR (conn.STATUS = 2);
END_FUNCTION_BLOCK

// Read DB bytes (RK512 FETCH) — covers FB_NLinkFetch.
FUNCTION_BLOCK FB_NLinkFetch
VAR_INPUT
    hLink : UDINT;               // from FB_NLinkOpen
    nArea : UDINT := 1;          // only eNLinkArea_DB (=1) is valid
    nDB : UDINT := 0;            // DB number 0..255
    nOffset : UDINT;             // byte offset in the DB, even, <=510
    nLen : UDINT;                // bytes, 1..510
    bExecute : BOOL;
    tTimeout : TIME := T#2S;
END_VAR
VAR_OUTPUT
    bBusy : BOOL;
    bDone : BOOL;
    bError : BOOL;
    nErrID : UDINT;
    nStatus : DINT;              // 0=pending 1=ok 2=timeout
                                  // 3=error 4=badresp 5=s5err
    cbRead : UDINT;              // bytes returned
    pBuffer : ARRAY[0..509] OF BYTE;
END_VAR
VAR
    io : FB_S5Io;
    i : UDINT;
END_VAR
    io.CONN_HANDLE := hLink;
    io.MODE := 0;
    io.DB := nDB;
    io.BYTE_OFF := nOffset;
    io.LEN := nLen;
    io.TIMEOUT := tTimeout;
    io.EXEC := bExecute;
    io();
    bBusy := io.BUSY;
    bDone := io.DONE;
    nStatus := io.STATUS;
    nErrID := io.ERRID;
    cbRead := io.DATA_LEN;
    IF io.DONE THEN
        i := 0;
        WHILE i < io.DATA_LEN AND i < 510 DO
            pBuffer[i] := io.R_DATA[i];
            i := i + 1;
        END_WHILE;
    END_IF;
    bError := (io.ERRID <> 0) OR (io.STATUS >= 2) OR (nArea <> 1);
END_FUNCTION_BLOCK

// Write DB bytes (RK512 SEND) — covers FB_NLinkWrite.
FUNCTION_BLOCK FB_NLinkWrite
VAR_INPUT
    hLink : UDINT;
    nArea : UDINT := 1;          // only eNLinkArea_DB (=1) is valid
    nDB : UDINT := 0;
    nOffset : UDINT;             // byte offset in the DB, even, <=510
    nLen : UDINT;                // bytes, 1..510
    pData : ARRAY[0..509] OF BYTE;
    bExecute : BOOL;
    tTimeout : TIME := T#2S;
END_VAR
VAR_OUTPUT
    bBusy : BOOL;
    bDone : BOOL;
    bError : BOOL;
    nErrID : UDINT;
    nStatus : DINT;
    cbWrite : UDINT;             // bytes accepted
END_VAR
VAR
    io : FB_S5Io;
    i : UDINT;
END_VAR
    io.CONN_HANDLE := hLink;
    io.MODE := 1;
    io.DB := nDB;
    io.BYTE_OFF := nOffset;
    io.LEN := nLen;
    io.TIMEOUT := tTimeout;
    i := 0;
    WHILE i < 510 DO
        io.DATA[i] := pData[i];
        i := i + 1;
    END_WHILE;
    io.EXEC := bExecute;
    io();
    bBusy := io.BUSY;
    bDone := io.DONE;
    nStatus := io.STATUS;
    nErrID := io.ERRID;
    cbWrite := 0;
    IF io.DONE AND io.STATUS = 1 THEN
        cbWrite := nLen;
    END_IF;
    bError := (io.ERRID <> 0) OR (io.STATUS >= 2) OR (nArea <> 1);
END_FUNCTION_BLOCK

// Library version query — covers F_GetVersionTcS5S7Comm.
FUNCTION F_GetVersionTcS5S7Comm : UINT
VAR_INPUT
    END_VAR
    F_GetVersionTcS5S7Comm := 16#0100;
END_FUNCTION

(* ---- tc2_serialcom.st ---- *)
// Tc2_SerialCom serial FBs (TwinCAT 3 PLC Library Tc2_SerialCom).
// Beckhoff-shaped wrappers over the builtin FB_Serial, which drives
// the host "tplc-serial" service (POSIX termios, nonblocking,
// deadline-bounded).
// TwinCAT's ComBuffer/SerialLineControl model keeps per-port state in
// a runtime-owned buffer object; this port uses explicit UDINT
// handles returned by FB_SerialOpen instead. Payload pointers
// (POINTER TO BYTE) are STRING[256] buffers.
// nParity: 0=none, 1=even, 2=odd. nStopBits: 1 or 2. nFlags is the
// TPLC_SERIAL_F_* bitmask (1=raw, 2=RS485, 4=noctty).
// Sources: docs/plc/plan/21-twincat-libraries.md §7 (TF6000).

FUNCTION_BLOCK FB_SerialOpen
VAR_INPUT
    bExecute : BOOL;
    tTimeout : TIME;
    sDevice : STRING[63];
    nBaud : UDINT;
    nParity : UDINT;
    nDataBits : UDINT;
    nStopBits : UDINT;
    nFlags : UDINT;
END_VAR
VAR_OUTPUT
    bBusy : BOOL;
    bDone : BOOL;
    bError : BOOL;
    nErrId : UDINT;
    hPort : UDINT;
END_VAR
VAR
    ser : FB_Serial;
END_VAR
    ser.OP := 1;
    ser.DEV := sDevice;
    ser.BAUD := nBaud;
    ser.PARITY := nParity;
    ser.DBITS := nDataBits;
    ser.SBITS := nStopBits;
    ser.FLAGS := nFlags;
    ser.TIMEOUT := tTimeout;
    ser.EXEC := bExecute;
    ser();
    bBusy := ser.BUSY;
    bDone := ser.DONE;
    nErrId := ser.ERRID;
    hPort := ser.HANDLE;
    bError := ser.ERRID <> 0;
END_FUNCTION_BLOCK

FUNCTION_BLOCK FB_SerialSend
VAR_INPUT
    bExecute : BOOL;
    tTimeout : TIME;
    hPort : UDINT;
    pData : STRING[256];
    nLen : UDINT;
END_VAR
VAR_OUTPUT
    bBusy : BOOL;
    bDone : BOOL;
    bError : BOOL;
    nErrId : UDINT;
    nSent : DINT;
END_VAR
VAR
    ser : FB_Serial;
END_VAR
    ser.OP := 2;
    ser.HANDLE := hPort;
    ser.DATA := pData;
    ser.DLEN := nLen;
    ser.TIMEOUT := tTimeout;
    ser.EXEC := bExecute;
    ser();
    bBusy := ser.BUSY;
    bDone := ser.DONE;
    nErrId := ser.ERRID;
    nSent := ser.RESULT;
    bError := ser.ERRID <> 0;
END_FUNCTION_BLOCK

FUNCTION_BLOCK FB_SerialReceive
VAR_INPUT
    bExecute : BOOL;
    tTimeout : TIME;
    hPort : UDINT;
END_VAR
VAR_OUTPUT
    bBusy : BOOL;
    bDone : BOOL;
    bError : BOOL;
    nErrId : UDINT;
    pData : STRING[256];
    nRecBytes : UDINT;
END_VAR
VAR
    ser : FB_Serial;
END_VAR
    ser.OP := 3;
    ser.HANDLE := hPort;
    ser.TIMEOUT := tTimeout;
    ser.EXEC := bExecute;
    ser();
    bBusy := ser.BUSY;
    bDone := ser.DONE;
    nErrId := ser.ERRID;
    pData := ser.DATA;
    nRecBytes := ser.DLEN;
    bError := ser.ERRID <> 0;
END_FUNCTION_BLOCK

FUNCTION_BLOCK FB_SerialClose
VAR_INPUT
    bExecute : BOOL;
    tTimeout : TIME;
    hPort : UDINT;
END_VAR
VAR_OUTPUT
    bBusy : BOOL;
    bDone : BOOL;
    bError : BOOL;
    nErrId : UDINT;
END_VAR
VAR
    ser : FB_Serial;
END_VAR
    ser.OP := 4;
    ser.HANDLE := hPort;
    ser.TIMEOUT := tTimeout;
    ser.EXEC := bExecute;
    ser();
    bBusy := ser.BUSY;
    bDone := ser.DONE;
    nErrId := ser.ERRID;
    bError := ser.ERRID <> 0;
END_FUNCTION_BLOCK

FUNCTION_BLOCK FB_SerialFlush
VAR_INPUT
    bExecute : BOOL;
    tTimeout : TIME;
    hPort : UDINT;
    nPurge : UDINT;
END_VAR
VAR_OUTPUT
    bBusy : BOOL;
    bDone : BOOL;
    bError : BOOL;
    nErrId : UDINT;
END_VAR
VAR
    ser : FB_Serial;
END_VAR
    ser.OP := 5;
    ser.HANDLE := hPort;
    ser.AUX := nPurge;
    ser.TIMEOUT := tTimeout;
    ser.EXEC := bExecute;
    ser();
    bBusy := ser.BUSY;
    bDone := ser.DONE;
    nErrId := ser.ERRID;
    bError := ser.ERRID <> 0;
END_FUNCTION_BLOCK

FUNCTION_BLOCK FB_SerialRs485
VAR_INPUT
    bExecute : BOOL;
    tTimeout : TIME;
    hPort : UDINT;
    bEnable : BOOL;
END_VAR
VAR_OUTPUT
    bBusy : BOOL;
    bDone : BOOL;
    bError : BOOL;
    nErrId : UDINT;
END_VAR
VAR
    ser : FB_Serial;
    en : UDINT;
END_VAR
    IF bEnable THEN
        en := 1;
    ELSE
        en := 0;
    END_IF
    ser.OP := 6;
    ser.HANDLE := hPort;
    ser.AUX := en;
    ser.TIMEOUT := tTimeout;
    ser.EXEC := bExecute;
    ser();
    bBusy := ser.BUSY;
    bDone := ser.DONE;
    nErrId := ser.ERRID;
    bError := ser.ERRID <> 0;
END_FUNCTION_BLOCK

(* ---- tc2_sms_sms.st ---- *)
// Tc2_SMS + Tc2_SMTP -> SMS-over-GSM-modem and SMTP client wrappers.
// TwinCAT's FB_Smtp* blocks proxy through a TwinCAT SMTP server
// over ADS; TetherPLC adapts them to a direct RFC 5321 client on
// the tplc-smtp service (poll model, one transaction per EXEC
// edge, plain text only, AUTH LOGIN when USER/PASS are set).
// SendSMS drives a GSM modem through the Tc2_SerialCom wrappers
// (tplc-serial service) with an AT-command state machine in text
// mode (AT+CMGF=1, AT+CMGS, SUB-terminated body).
// Differences from the TwinCAT blocks, documented in
// docs/plc/compat/README.md:
//   - No ADS SMTP server proxy, no TLS/SSL, no attachments
//     (FB_SmtpAttach reports an unsupported error), no delivery
//     receipts, no multi-recipient envelopes (single RCPT TO),
//     no MIME headers beyond Subject/From/To/Date.
//   - SMS: PDU mode, concatenated SMS (UCS2), status reports and
//     delivery reports are not implemented; the modem must
//     support AT+CMGF=1 text mode. sText is limited to 160 chars
//     (one GSM-7 segment); longer texts are truncated by the
//     serial channel.
// Sources: docs/plc/plan/21-twincat-libraries.md (TF6350 SMS/SMTP).

// SMTP send without authentication — TwinCAT FB_SmtpV3 subset.
// nStatus mirrors TplcSmtpInfo: 0=pending 1=ok 2=fail(smtp reply
// code in nRespCode) 3=timeout 4=error 5=badresp.
FUNCTION_BLOCK FB_SmtpV3
VAR_INPUT
    bExecute : BOOL;
    tTimeout : TIME := T#10S;
    sServer : STRING[15];          // dotted-quad IPv4
    nPort : UDINT := 25;           // 0 = 25
    sFrom : STRING[63];
    sTo : STRING[63];
    sSubject : STRING[63];
    sBody : STRING[255];
END_VAR
VAR_OUTPUT
    bBusy : BOOL;
    bDone : BOOL;
    bError : BOOL;
    nErrId : UDINT;
    nStatus : DINT;
    nRespCode : UDINT;
END_VAR
VAR
    smtp : FB_SmtpSend;
END_VAR
    smtp.HOST := sServer;
    smtp.PORT := nPort;
    smtp.USER := '';
    smtp.PASS := '';
    smtp.FROM := sFrom;
    smtp.RCPT := sTo;
    smtp.SUBJECT := sSubject;
    smtp.TIMEOUT := tTimeout;
    smtp.BODY := sBody;
    smtp.EXEC := bExecute;
    smtp();
    bBusy := smtp.BUSY;
    bDone := smtp.DONE;
    nStatus := smtp.STATUS;
    nRespCode := smtp.RESP_CODE;
    nErrId := smtp.ERRID;
    bError := smtp.BUSY = FALSE AND smtp.DONE = TRUE AND smtp.STATUS >= 2;
END_FUNCTION_BLOCK

// SMTP send with AUTH LOGIN — TwinCAT FB_SmtpV3_Full subset.
// sUser/sPass empty disables authentication (same as FB_SmtpV3).
FUNCTION_BLOCK FB_SmtpV3_Full
VAR_INPUT
    bExecute : BOOL;
    tTimeout : TIME := T#10S;
    sServer : STRING[15];
    nPort : UDINT := 25;
    sUser : STRING[31];
    sPass : STRING[31];
    sFrom : STRING[63];
    sTo : STRING[63];
    sSubject : STRING[63];
    sBody : STRING[255];
END_VAR
VAR_OUTPUT
    bBusy : BOOL;
    bDone : BOOL;
    bError : BOOL;
    nErrId : UDINT;
    nStatus : DINT;
    nRespCode : UDINT;
END_VAR
VAR
    smtp : FB_SmtpSend;
END_VAR
    smtp.HOST := sServer;
    smtp.PORT := nPort;
    smtp.USER := sUser;
    smtp.PASS := sPass;
    smtp.FROM := sFrom;
    smtp.RCPT := sTo;
    smtp.SUBJECT := sSubject;
    smtp.TIMEOUT := tTimeout;
    smtp.BODY := sBody;
    smtp.EXEC := bExecute;
    smtp();
    bBusy := smtp.BUSY;
    bDone := smtp.DONE;
    nStatus := smtp.STATUS;
    nRespCode := smtp.RESP_CODE;
    nErrId := smtp.ERRID;
    bError := smtp.BUSY = FALSE AND smtp.DONE = TRUE AND smtp.STATUS >= 2;
END_FUNCTION_BLOCK

// Obsolete TwinCAT FB_Smtp — kept as an alias of FB_SmtpV3.
FUNCTION_BLOCK FB_Smtp
VAR_INPUT
    bExecute : BOOL;
    tTimeout : TIME := T#10S;
    sServer : STRING[15];
    nPort : UDINT := 25;
    sFrom : STRING[63];
    sTo : STRING[63];
    sSubject : STRING[63];
    sBody : STRING[255];
END_VAR
VAR_OUTPUT
    bBusy : BOOL;
    bDone : BOOL;
    bError : BOOL;
    nErrId : UDINT;
    nStatus : DINT;
    nRespCode : UDINT;
END_VAR
VAR
    v3 : FB_SmtpV3;
END_VAR
    v3.bExecute := bExecute;
    v3.tTimeout := tTimeout;
    v3.sServer := sServer;
    v3.nPort := nPort;
    v3.sFrom := sFrom;
    v3.sTo := sTo;
    v3.sSubject := sSubject;
    v3.sBody := sBody;
    v3();
    bBusy := v3.bBusy;
    bDone := v3.bDone;
    bError := v3.bError;
    nErrId := v3.nErrId;
    nStatus := v3.nStatus;
    nRespCode := v3.nRespCode;
END_FUNCTION_BLOCK

// Obsolete TwinCAT FB_SmtpFull — alias of FB_SmtpV3_Full.
FUNCTION_BLOCK FB_SmtpFull
VAR_INPUT
    bExecute : BOOL;
    tTimeout : TIME := T#10S;
    sServer : STRING[15];
    nPort : UDINT := 25;
    sUser : STRING[31];
    sPass : STRING[31];
    sFrom : STRING[63];
    sTo : STRING[63];
    sSubject : STRING[63];
    sBody : STRING[255];
END_VAR
VAR_OUTPUT
    bBusy : BOOL;
    bDone : BOOL;
    bError : BOOL;
    nErrId : UDINT;
    nStatus : DINT;
    nRespCode : UDINT;
END_VAR
VAR
    v3 : FB_SmtpV3_Full;
END_VAR
    v3.bExecute := bExecute;
    v3.tTimeout := tTimeout;
    v3.sServer := sServer;
    v3.nPort := nPort;
    v3.sUser := sUser;
    v3.sPass := sPass;
    v3.sFrom := sFrom;
    v3.sTo := sTo;
    v3.sSubject := sSubject;
    v3.sBody := sBody;
    v3();
    bBusy := v3.bBusy;
    bDone := v3.bDone;
    bError := v3.bError;
    nErrId := v3.nErrId;
    nStatus := v3.nStatus;
    nRespCode := v3.nRespCode;
END_FUNCTION_BLOCK

// TwinCAT FB_SmtpAttach — MIME file attachment. TetherPLC has no
// MIME/base64 encoder in the ST layer, so this FB reports an
// unsupported error immediately on EXEC. nErrId = 90.
FUNCTION_BLOCK FB_SmtpAttach
VAR_INPUT
    bExecute : BOOL;
    tTimeout : TIME := T#10S;
    sServer : STRING[15];
    nPort : UDINT := 25;
    sUser : STRING[31];
    sPass : STRING[31];
    sFrom : STRING[63];
    sTo : STRING[63];
    sSubject : STRING[63];
    sBody : STRING[255];
    sAttachPath : STRING[63];
END_VAR
VAR_OUTPUT
    bBusy : BOOL;
    bDone : BOOL;
    bError : BOOL;
    nErrId : UDINT;
    nStatus : DINT;
    nRespCode : UDINT;
END_VAR
VAR
    lastExec : BOOL;
END_VAR
    IF bExecute AND NOT lastExec THEN
        bBusy := FALSE;
        bDone := TRUE;
        bError := TRUE;
        nErrId := 90;
        nStatus := 4;
        nRespCode := 0;
    ELSE
        bBusy := FALSE;
        bDone := FALSE;
        bError := FALSE;
        nErrId := 0;
        nStatus := 0;
        nRespCode := 0;
    END_IF;
    lastExec := bExecute;
END_FUNCTION_BLOCK

// GSM SMS send — TwinCAT SendSMS adapted to the poll model.
// hPort is an open serial handle from FB_SerialOpen (the modem
// UART). The FB runs the AT sequence autonomously after a
// rising edge on bExecute:
//   AT -> AT+CMGF=1 -> AT+CMGS="<sNumber>" -> sText + SUB(0x1A)
// nStatus: 0=ok 1=timeout 2=modem error 3=serial error.
// sLastRx keeps the tail of the modem response for diagnostics.
FUNCTION_BLOCK FB_SendSMS
VAR_INPUT
    bExecute : BOOL;
    tTimeout : TIME := T#10S;   // per-command budget hint
    hPort : UDINT;              // open handle from FB_SerialOpen
    sNumber : STRING[31];       // destination number
    sText : STRING[160];        // GSM-7 text, 160 chars max
END_VAR
VAR_OUTPUT
    bBusy : BOOL;
    bDone : BOOL;
    bError : BOOL;
    nErrId : UDINT;
    nStatus : DINT;
    sLastRx : STRING[255];
    dbgPhase : INT;
    dbgTries : UDINT;
END_VAR
VAR
    st : INT;
    phase : INT;                // 0=send cmd 1=await reply
    tries : UDINT;
    cmd : STRING[256];
    tokOk : STRING[8];
    tokOk2 : STRING[8];
    tokErr : STRING[8];
    rxAcc : STRING[512];
    ctrlZ : STRING[1];
    lastExec : BOOL;
    snd : FB_SerialSend;
    rcv : FB_SerialReceive;
    sndKick : BOOL;
    rcvKick : BOOL;
END_VAR

    IF bExecute AND NOT lastExec AND st = 0 THEN
        st := 1;
        phase := 0;
        tries := 0;
        rxAcc := '';
        ctrlZ := '';
        cmd := 'AT$R';
        tokOk := 'OK';
        tokOk2 := '';
        tokErr := '';
        sndKick := TRUE;
    END_IF;
    lastExec := bExecute;

    // Both serial FBs are called every scan with bExecute pulsed
    // only on kick scans. FB_Serial arms on a 0->1 EXEC edge, so
    // EXEC must see a low scan between transactions; gating the
    // calls by phase would freeze EXEC high after a fast write
    // and swallow the next kick.
    snd.bExecute := sndKick AND (phase = 0);
    sndKick := FALSE;
    snd.tTimeout := T#2S;
    snd.hPort := hPort;
    snd.pData := cmd;
    snd.nLen := 0;
    snd();

    rcv.bExecute := rcvKick AND (phase = 1);
    rcvKick := FALSE;
    rcv.tTimeout := T#400MS;
    rcv.hPort := hPort;
    rcv();

    IF st >= 1 AND st <= 4 THEN
        IF phase = 0 AND snd.bDone THEN
            IF snd.nErrId <> 0 THEN
                st := 9;
                nStatus := 3;
                nErrId := snd.nErrId;
            ELSE
                phase := 1;
                tries := 0;
                rxAcc := '';
                rcvKick := TRUE;
            END_IF;
        ELSIF phase = 1 AND rcv.bDone THEN
            // await leg: each read completion appends to rxAcc
            // and rescans for the expected token. ~25 x 400ms.
                IF rcv.nErrId = 0 AND rcv.nRecBytes > 0 THEN
                    IF LEN(rxAcc) > 200 THEN
                        st := 9;
                        nStatus := 2;
                        nErrId := 91;
                    ELSE
                        rxAcc := CONCAT(rxAcc, rcv.pData);
                        sLastRx := rcv.pData;
                        IF tokErr <> '' AND FIND(rxAcc, tokErr) > 0 THEN
                            st := 9;
                            nStatus := 2;
                            nErrId := 92;
                        ELSIF FIND(rxAcc, tokOk) > 0
                            OR (tokOk2 <> '' AND FIND(rxAcc, tokOk2) > 0) THEN
                            IF st = 1 THEN
                                st := 2; phase := 0; sndKick := TRUE;
                                cmd := 'AT+CMGF=1$R';
                                tokOk := 'OK'; tokOk2 := '';
                            ELSIF st = 2 THEN
                                st := 3; phase := 0; sndKick := TRUE;
                                cmd := CONCAT('AT+CMGS="', sNumber);
                                cmd := CONCAT(cmd, '"$R');
                                tokOk := '>'; tokOk2 := '';
                            ELSIF st = 3 THEN
                                st := 4; phase := 0; sndKick := TRUE;
                                cmd := CONCAT(sText, ctrlZ);
                                tokOk := '+CMGS'; tokOk2 := 'OK';
                                tokErr := 'ERROR';
                            ELSE
                                st := 5;
                            END_IF;
                            tries := 0;
                            rxAcc := '';
                        ELSE
                            tries := tries + 1;
                            IF tries > 25 THEN
                                st := 9;
                                nStatus := 1;
                                nErrId := 5;
                            ELSE
                                rcvKick := TRUE;
                            END_IF;
                        END_IF;
                    END_IF;
                ELSE
                    tries := tries + 1;
                    IF tries > 25 THEN
                        st := 9;
                        nStatus := 1;
                        nErrId := 5;
                    ELSE
                        rcvKick := TRUE;
                    END_IF;
                END_IF;
        END_IF;
        bBusy := TRUE;
        bDone := FALSE;
        bError := FALSE;
        dbgPhase := st * 10 + phase;
        dbgTries := tries;
    ELSIF st = 5 THEN
        bBusy := FALSE;
        bDone := TRUE;
        bError := FALSE;
        nStatus := 0;
        nErrId := 0;
        st := 6;
    ELSIF st = 6 THEN
        bBusy := FALSE;
        bDone := FALSE;
        bError := FALSE;
        nStatus := 0;
        nErrId := 0;
        st := 0;
    ELSIF st = 9 THEN
        bBusy := FALSE;
        bDone := TRUE;
        bError := TRUE;
        st := 10;
    ELSIF st = 10 THEN
        bBusy := FALSE;
        bDone := FALSE;
        bError := FALSE;
        st := 0;
    ELSE
        bBusy := FALSE;
        bDone := FALSE;
        bError := FALSE;
        nStatus := 0;
        nErrId := 0;
    END_IF;
END_FUNCTION_BLOCK

// TwinCAT Get_TcPlcSMS_Version — returns the SMS layer version
// string after one EXEC edge. sVersion is fixed; nErrId = 0.
FUNCTION_BLOCK FB_GetTcPlcSMS_Version
VAR_INPUT
    bExecute : BOOL;
END_VAR
VAR_OUTPUT
    bBusy : BOOL;
    bDone : BOOL;
    sVersion : STRING[31];
END_VAR
VAR
    lastExec : BOOL;
    fired : BOOL;
END_VAR
    IF bExecute AND NOT lastExec AND NOT fired THEN
        fired := TRUE;
        sVersion := 'TetherPLC-TcSMS 1.0';
    END_IF;
    lastExec := bExecute;
    bBusy := FALSE;
    bDone := fired;
END_FUNCTION_BLOCK
